(* IEC 61131-3 sources: 2026_Projet_YGO_ExcavatriceDragage/TOOLS/TEST_AUTO_CI/RESULTS/L_SIMULATION/tests (part 8) *)

TEST 'TC-T418-INT-004 Premier geste N2 observe HX1 existant'
nx := 5000; ny := 5000; raw1 := 0; raw2 := 0; previousButton := FALSE; buttonEdges := 0;
bench.Enable := TRUE; joy.Enable := TRUE; joy.ArmingPermit := TRUE; diagOk.Operational := TRUE;
joy.BusCanOpenOP := diagOk; joy.JoystickOP := diagOk; home.Enable := TRUE; home.BootReady := TRUE;
home.Mode := E_Mode.MAINT_N2; home.BucketOffsetValid := TRUE; home.WinchesMechanicallyStopped := TRUE;
ADVANCE_TIME(10000000);
bench(RawPosM1 := raw1, RawPosM2 := raw2);
joy(RawX := bench.Operator.JoyXRaw_ANA1, RawY := bench.Operator.JoyYRaw_ANA2, RawButton := bench.Operator.JoyBtnRaw, Cfg := cfg, NeutralXMem := nx, NeutralYMem := ny);
home(DeadmanArmed := joy.DeadmanArmed, JoystickDeflected := NOT joy.AtNeutralXY, JoystickPull := joy.AxisCmdY.DirectionPositive, JoystickPush := joy.AxisCmdY.DirectionNegative, BtnValidation := bench.Operator.JoyBtnRaw);
IF bench.Operator.JoyBtnRaw AND NOT previousButton THEN buttonEdges := buttonEdges + 1; END_IF; previousButton := bench.Operator.JoyBtnRaw;
bench.SimJoystickRight_Fwd_MAINT_Active := TRUE;
ADVANCE_TIME(10000000);
bench(RawPosM1 := raw1, RawPosM2 := raw2);
joy(RawX := bench.Operator.JoyXRaw_ANA1, RawY := bench.Operator.JoyYRaw_ANA2, RawButton := bench.Operator.JoyBtnRaw, Cfg := cfg, NeutralXMem := nx, NeutralYMem := ny);
home(DeadmanArmed := joy.DeadmanArmed, JoystickDeflected := NOT joy.AtNeutralXY, JoystickPull := joy.AxisCmdY.DirectionPositive, JoystickPush := joy.AxisCmdY.DirectionNegative, BtnValidation := bench.Operator.JoyBtnRaw);
IF bench.Operator.JoyBtnRaw AND NOT previousButton THEN buttonEdges := buttonEdges + 1; END_IF; previousButton := bench.Operator.JoyBtnRaw;
ASSERT_EQ(home.MachineHomingSeqStep, E_MachineHomingTxState.HX1_BUCKET_PREPARE, 'CONSTAT production : front homme-mort lance HX1 en N2');
ADVANCE_TIME(10000000);
bench(RawPosM1 := raw1, RawPosM2 := raw2);
joy(RawX := bench.Operator.JoyXRaw_ANA1, RawY := bench.Operator.JoyYRaw_ANA2, RawButton := bench.Operator.JoyBtnRaw, Cfg := cfg, NeutralXMem := nx, NeutralYMem := ny);
home(DeadmanArmed := joy.DeadmanArmed, JoystickDeflected := NOT joy.AtNeutralXY, JoystickPull := joy.AxisCmdY.DirectionPositive, JoystickPush := joy.AxisCmdY.DirectionNegative, BtnValidation := bench.Operator.JoyBtnRaw);
IF bench.Operator.JoyBtnRaw AND NOT previousButton THEN buttonEdges := buttonEdges + 1; END_IF; previousButton := bench.Operator.JoyBtnRaw;
ASSERT_TRUE(home.M3Locked, 'CONSTAT production : homing verrouille M3'); ASSERT_EQ(buttonEdges, 1, 'Front fidele non masque');
END_TEST

TEST 'TC-T418-INT-005 Stimuli manuels exclusifs et pas de saut au retour'
nx := 5000; ny := 5000; raw1 := 0; raw2 := 0; previousButton := FALSE; buttonEdges := 0;
bench.Enable := TRUE; joy.Enable := TRUE; joy.ArmingPermit := TRUE; diagOk.Operational := TRUE;
joy.BusCanOpenOP := diagOk; joy.JoystickOP := diagOk; home.Enable := TRUE; home.BootReady := TRUE;
home.Mode := E_Mode.MAINT_N1; home.BucketOffsetValid := TRUE; home.WinchesMechanicallyStopped := TRUE;
ADVANCE_TIME(10000000);
bench(RawPosM1 := raw1, RawPosM2 := raw2);
joy(RawX := bench.Operator.JoyXRaw_ANA1, RawY := bench.Operator.JoyYRaw_ANA2, RawButton := bench.Operator.JoyBtnRaw, Cfg := cfg, NeutralXMem := nx, NeutralYMem := ny);
home(DeadmanArmed := joy.DeadmanArmed, JoystickDeflected := NOT joy.AtNeutralXY, JoystickPull := joy.AxisCmdY.DirectionPositive, JoystickPush := joy.AxisCmdY.DirectionNegative, BtnValidation := bench.Operator.JoyBtnRaw);
IF bench.Operator.JoyBtnRaw AND NOT previousButton THEN buttonEdges := buttonEdges + 1; END_IF; previousButton := bench.Operator.JoyBtnRaw;
bench.SimJoystickRawX := 8000; bench.SimJoystickRawButton := TRUE;
ADVANCE_TIME(10000000);
bench(RawPosM1 := raw1, RawPosM2 := raw2);
joy(RawX := bench.Operator.JoyXRaw_ANA1, RawY := bench.Operator.JoyYRaw_ANA2, RawButton := bench.Operator.JoyBtnRaw, Cfg := cfg, NeutralXMem := nx, NeutralYMem := ny);
home(DeadmanArmed := joy.DeadmanArmed, JoystickDeflected := NOT joy.AtNeutralXY, JoystickPull := joy.AxisCmdY.DirectionPositive, JoystickPush := joy.AxisCmdY.DirectionNegative, BtnValidation := bench.Operator.JoyBtnRaw);
IF bench.Operator.JoyBtnRaw AND NOT previousButton THEN buttonEdges := buttonEdges + 1; END_IF; previousButton := bench.Operator.JoyBtnRaw;
ASSERT_EQ(bench.Operator.JoyXRaw_ANA1, 8000, 'Manuel disponible au repos'); ASSERT_TRUE(bench.Operator.JoyBtnRaw, 'Bouton manuel publie');
bench.SimJoystickRight_Fwd_MAINT_Active := TRUE;
ADVANCE_TIME(10000000);
bench(RawPosM1 := raw1, RawPosM2 := raw2);
joy(RawX := bench.Operator.JoyXRaw_ANA1, RawY := bench.Operator.JoyYRaw_ANA2, RawButton := bench.Operator.JoyBtnRaw, Cfg := cfg, NeutralXMem := nx, NeutralYMem := ny);
home(DeadmanArmed := joy.DeadmanArmed, JoystickDeflected := NOT joy.AtNeutralXY, JoystickPull := joy.AxisCmdY.DirectionPositive, JoystickPush := joy.AxisCmdY.DirectionNegative, BtnValidation := bench.Operator.JoyBtnRaw);
IF bench.Operator.JoyBtnRaw AND NOT previousButton THEN buttonEdges := buttonEdges + 1; END_IF; previousButton := bench.Operator.JoyBtnRaw;
ADVANCE_TIME(10000000);
bench(RawPosM1 := raw1, RawPosM2 := raw2);
joy(RawX := bench.Operator.JoyXRaw_ANA1, RawY := bench.Operator.JoyYRaw_ANA2, RawButton := bench.Operator.JoyBtnRaw, Cfg := cfg, NeutralXMem := nx, NeutralYMem := ny);
home(DeadmanArmed := joy.DeadmanArmed, JoystickDeflected := NOT joy.AtNeutralXY, JoystickPull := joy.AxisCmdY.DirectionPositive, JoystickPush := joy.AxisCmdY.DirectionNegative, BtnValidation := bench.Operator.JoyBtnRaw);
IF bench.Operator.JoyBtnRaw AND NOT previousButton THEN buttonEdges := buttonEdges + 1; END_IF; previousButton := bench.Operator.JoyBtnRaw;
ADVANCE_TIME(10000000);
bench(RawPosM1 := raw1, RawPosM2 := raw2);
joy(RawX := bench.Operator.JoyXRaw_ANA1, RawY := bench.Operator.JoyYRaw_ANA2, RawButton := bench.Operator.JoyBtnRaw, Cfg := cfg, NeutralXMem := nx, NeutralYMem := ny);
home(DeadmanArmed := joy.DeadmanArmed, JoystickDeflected := NOT joy.AtNeutralXY, JoystickPull := joy.AxisCmdY.DirectionPositive, JoystickPush := joy.AxisCmdY.DirectionNegative, BtnValidation := bench.Operator.JoyBtnRaw);
IF bench.Operator.JoyBtnRaw AND NOT previousButton THEN buttonEdges := buttonEdges + 1; END_IF; previousButton := bench.Operator.JoyBtnRaw;
ADVANCE_TIME(10000000);
bench(RawPosM1 := raw1, RawPosM2 := raw2);
joy(RawX := bench.Operator.JoyXRaw_ANA1, RawY := bench.Operator.JoyYRaw_ANA2, RawButton := bench.Operator.JoyBtnRaw, Cfg := cfg, NeutralXMem := nx, NeutralYMem := ny);
home(DeadmanArmed := joy.DeadmanArmed, JoystickDeflected := NOT joy.AtNeutralXY, JoystickPull := joy.AxisCmdY.DirectionPositive, JoystickPush := joy.AxisCmdY.DirectionNegative, BtnValidation := bench.Operator.JoyBtnRaw);
IF bench.Operator.JoyBtnRaw AND NOT previousButton THEN buttonEdges := buttonEdges + 1; END_IF; previousButton := bench.Operator.JoyBtnRaw;
ADVANCE_TIME(10000000);
bench(RawPosM1 := raw1, RawPosM2 := raw2);
joy(RawX := bench.Operator.JoyXRaw_ANA1, RawY := bench.Operator.JoyYRaw_ANA2, RawButton := bench.Operator.JoyBtnRaw, Cfg := cfg, NeutralXMem := nx, NeutralYMem := ny);
home(DeadmanArmed := joy.DeadmanArmed, JoystickDeflected := NOT joy.AtNeutralXY, JoystickPull := joy.AxisCmdY.DirectionPositive, JoystickPush := joy.AxisCmdY.DirectionNegative, BtnValidation := bench.Operator.JoyBtnRaw);
IF bench.Operator.JoyBtnRaw AND NOT previousButton THEN buttonEdges := buttonEdges + 1; END_IF; previousButton := bench.Operator.JoyBtnRaw;
ASSERT_EQ(bench.Operator.JoyXRaw_ANA1, 5000, 'Conflit manuel automatique neutralise'); ASSERT_FALSE(bench.Operator.JoyBtnRaw, 'Aucun OR des sources');
bench.SimJoystickRawX := 5000; bench.SimJoystickRawButton := FALSE;
ADVANCE_TIME(10000000);
bench(RawPosM1 := raw1, RawPosM2 := raw2);
joy(RawX := bench.Operator.JoyXRaw_ANA1, RawY := bench.Operator.JoyYRaw_ANA2, RawButton := bench.Operator.JoyBtnRaw, Cfg := cfg, NeutralXMem := nx, NeutralYMem := ny);
home(DeadmanArmed := joy.DeadmanArmed, JoystickDeflected := NOT joy.AtNeutralXY, JoystickPull := joy.AxisCmdY.DirectionPositive, JoystickPush := joy.AxisCmdY.DirectionNegative, BtnValidation := bench.Operator.JoyBtnRaw);
IF bench.Operator.JoyBtnRaw AND NOT previousButton THEN buttonEdges := buttonEdges + 1; END_IF; previousButton := bench.Operator.JoyBtnRaw;
ADVANCE_TIME(10000000);
bench(RawPosM1 := raw1, RawPosM2 := raw2);
joy(RawX := bench.Operator.JoyXRaw_ANA1, RawY := bench.Operator.JoyYRaw_ANA2, RawButton := bench.Operator.JoyBtnRaw, Cfg := cfg, NeutralXMem := nx, NeutralYMem := ny);
home(DeadmanArmed := joy.DeadmanArmed, JoystickDeflected := NOT joy.AtNeutralXY, JoystickPull := joy.AxisCmdY.DirectionPositive, JoystickPush := joy.AxisCmdY.DirectionNegative, BtnValidation := bench.Operator.JoyBtnRaw);
IF bench.Operator.JoyBtnRaw AND NOT previousButton THEN buttonEdges := buttonEdges + 1; END_IF; previousButton := bench.Operator.JoyBtnRaw;
ADVANCE_TIME(10000000);
bench(RawPosM1 := raw1, RawPosM2 := raw2);
joy(RawX := bench.Operator.JoyXRaw_ANA1, RawY := bench.Operator.JoyYRaw_ANA2, RawButton := bench.Operator.JoyBtnRaw, Cfg := cfg, NeutralXMem := nx, NeutralYMem := ny);
home(DeadmanArmed := joy.DeadmanArmed, JoystickDeflected := NOT joy.AtNeutralXY, JoystickPull := joy.AxisCmdY.DirectionPositive, JoystickPush := joy.AxisCmdY.DirectionNegative, BtnValidation := bench.Operator.JoyBtnRaw);
IF bench.Operator.JoyBtnRaw AND NOT previousButton THEN buttonEdges := buttonEdges + 1; END_IF; previousButton := bench.Operator.JoyBtnRaw;
ADVANCE_TIME(10000000);
bench(RawPosM1 := raw1, RawPosM2 := raw2);
joy(RawX := bench.Operator.JoyXRaw_ANA1, RawY := bench.Operator.JoyYRaw_ANA2, RawButton := bench.Operator.JoyBtnRaw, Cfg := cfg, NeutralXMem := nx, NeutralYMem := ny);
home(DeadmanArmed := joy.DeadmanArmed, JoystickDeflected := NOT joy.AtNeutralXY, JoystickPull := joy.AxisCmdY.DirectionPositive, JoystickPush := joy.AxisCmdY.DirectionNegative, BtnValidation := bench.Operator.JoyBtnRaw);
IF bench.Operator.JoyBtnRaw AND NOT previousButton THEN buttonEdges := buttonEdges + 1; END_IF; previousButton := bench.Operator.JoyBtnRaw;
ADVANCE_TIME(10000000);
bench(RawPosM1 := raw1, RawPosM2 := raw2);
joy(RawX := bench.Operator.JoyXRaw_ANA1, RawY := bench.Operator.JoyYRaw_ANA2, RawButton := bench.Operator.JoyBtnRaw, Cfg := cfg, NeutralXMem := nx, NeutralYMem := ny);
home(DeadmanArmed := joy.DeadmanArmed, JoystickDeflected := NOT joy.AtNeutralXY, JoystickPull := joy.AxisCmdY.DirectionPositive, JoystickPush := joy.AxisCmdY.DirectionNegative, BtnValidation := bench.Operator.JoyBtnRaw);
IF bench.Operator.JoyBtnRaw AND NOT previousButton THEN buttonEdges := buttonEdges + 1; END_IF; previousButton := bench.Operator.JoyBtnRaw;
ASSERT_FALSE(bench.Operator.JoyBtnRaw, 'Enlever stimulus ne demarre pas bouton tenu');
bench.SimJoystickRight_Fwd_MAINT_Active := FALSE;
ADVANCE_TIME(10000000);
bench(RawPosM1 := raw1, RawPosM2 := raw2);
joy(RawX := bench.Operator.JoyXRaw_ANA1, RawY := bench.Operator.JoyYRaw_ANA2, RawButton := bench.Operator.JoyBtnRaw, Cfg := cfg, NeutralXMem := nx, NeutralYMem := ny);
home(DeadmanArmed := joy.DeadmanArmed, JoystickDeflected := NOT joy.AtNeutralXY, JoystickPull := joy.AxisCmdY.DirectionPositive, JoystickPush := joy.AxisCmdY.DirectionNegative, BtnValidation := bench.Operator.JoyBtnRaw);
IF bench.Operator.JoyBtnRaw AND NOT previousButton THEN buttonEdges := buttonEdges + 1; END_IF; previousButton := bench.Operator.JoyBtnRaw;
bench.SimJoystickRight_Fwd_MAINT_Active := TRUE;
ADVANCE_TIME(10000000);
bench(RawPosM1 := raw1, RawPosM2 := raw2);
joy(RawX := bench.Operator.JoyXRaw_ANA1, RawY := bench.Operator.JoyYRaw_ANA2, RawButton := bench.Operator.JoyBtnRaw, Cfg := cfg, NeutralXMem := nx, NeutralYMem := ny);
home(DeadmanArmed := joy.DeadmanArmed, JoystickDeflected := NOT joy.AtNeutralXY, JoystickPull := joy.AxisCmdY.DirectionPositive, JoystickPush := joy.AxisCmdY.DirectionNegative, BtnValidation := bench.Operator.JoyBtnRaw);
IF bench.Operator.JoyBtnRaw AND NOT previousButton THEN buttonEdges := buttonEdges + 1; END_IF; previousButton := bench.Operator.JoyBtnRaw;
ADVANCE_TIME(10000000);
bench(RawPosM1 := raw1, RawPosM2 := raw2);
joy(RawX := bench.Operator.JoyXRaw_ANA1, RawY := bench.Operator.JoyYRaw_ANA2, RawButton := bench.Operator.JoyBtnRaw, Cfg := cfg, NeutralXMem := nx, NeutralYMem := ny);
home(DeadmanArmed := joy.DeadmanArmed, JoystickDeflected := NOT joy.AtNeutralXY, JoystickPull := joy.AxisCmdY.DirectionPositive, JoystickPush := joy.AxisCmdY.DirectionNegative, BtnValidation := bench.Operator.JoyBtnRaw);
IF bench.Operator.JoyBtnRaw AND NOT previousButton THEN buttonEdges := buttonEdges + 1; END_IF; previousButton := bench.Operator.JoyBtnRaw;
ADVANCE_TIME(10000000);
bench(RawPosM1 := raw1, RawPosM2 := raw2);
joy(RawX := bench.Operator.JoyXRaw_ANA1, RawY := bench.Operator.JoyYRaw_ANA2, RawButton := bench.Operator.JoyBtnRaw, Cfg := cfg, NeutralXMem := nx, NeutralYMem := ny);
home(DeadmanArmed := joy.DeadmanArmed, JoystickDeflected := NOT joy.AtNeutralXY, JoystickPull := joy.AxisCmdY.DirectionPositive, JoystickPush := joy.AxisCmdY.DirectionNegative, BtnValidation := bench.Operator.JoyBtnRaw);
IF bench.Operator.JoyBtnRaw AND NOT previousButton THEN buttonEdges := buttonEdges + 1; END_IF; previousButton := bench.Operator.JoyBtnRaw;
ADVANCE_TIME(10000000);
bench(RawPosM1 := raw1, RawPosM2 := raw2);
joy(RawX := bench.Operator.JoyXRaw_ANA1, RawY := bench.Operator.JoyYRaw_ANA2, RawButton := bench.Operator.JoyBtnRaw, Cfg := cfg, NeutralXMem := nx, NeutralYMem := ny);
home(DeadmanArmed := joy.DeadmanArmed, JoystickDeflected := NOT joy.AtNeutralXY, JoystickPull := joy.AxisCmdY.DirectionPositive, JoystickPush := joy.AxisCmdY.DirectionNegative, BtnValidation := bench.Operator.JoyBtnRaw);
IF bench.Operator.JoyBtnRaw AND NOT previousButton THEN buttonEdges := buttonEdges + 1; END_IF; previousButton := bench.Operator.JoyBtnRaw;
ADVANCE_TIME(10000000);
bench(RawPosM1 := raw1, RawPosM2 := raw2);
joy(RawX := bench.Operator.JoyXRaw_ANA1, RawY := bench.Operator.JoyYRaw_ANA2, RawButton := bench.Operator.JoyBtnRaw, Cfg := cfg, NeutralXMem := nx, NeutralYMem := ny);
home(DeadmanArmed := joy.DeadmanArmed, JoystickDeflected := NOT joy.AtNeutralXY, JoystickPull := joy.AxisCmdY.DirectionPositive, JoystickPush := joy.AxisCmdY.DirectionNegative, BtnValidation := bench.Operator.JoyBtnRaw);
IF bench.Operator.JoyBtnRaw AND NOT previousButton THEN buttonEdges := buttonEdges + 1; END_IF; previousButton := bench.Operator.JoyBtnRaw;
ADVANCE_TIME(10000000);
bench(RawPosM1 := raw1, RawPosM2 := raw2);
joy(RawX := bench.Operator.JoyXRaw_ANA1, RawY := bench.Operator.JoyYRaw_ANA2, RawButton := bench.Operator.JoyBtnRaw, Cfg := cfg, NeutralXMem := nx, NeutralYMem := ny);
home(DeadmanArmed := joy.DeadmanArmed, JoystickDeflected := NOT joy.AtNeutralXY, JoystickPull := joy.AxisCmdY.DirectionPositive, JoystickPush := joy.AxisCmdY.DirectionNegative, BtnValidation := bench.Operator.JoyBtnRaw);
IF bench.Operator.JoyBtnRaw AND NOT previousButton THEN buttonEdges := buttonEdges + 1; END_IF; previousButton := bench.Operator.JoyBtnRaw;
ADVANCE_TIME(10000000);
bench(RawPosM1 := raw1, RawPosM2 := raw2);
joy(RawX := bench.Operator.JoyXRaw_ANA1, RawY := bench.Operator.JoyYRaw_ANA2, RawButton := bench.Operator.JoyBtnRaw, Cfg := cfg, NeutralXMem := nx, NeutralYMem := ny);
home(DeadmanArmed := joy.DeadmanArmed, JoystickDeflected := NOT joy.AtNeutralXY, JoystickPull := joy.AxisCmdY.DirectionPositive, JoystickPush := joy.AxisCmdY.DirectionNegative, BtnValidation := bench.Operator.JoyBtnRaw);
IF bench.Operator.JoyBtnRaw AND NOT previousButton THEN buttonEdges := buttonEdges + 1; END_IF; previousButton := bench.Operator.JoyBtnRaw;
ADVANCE_TIME(10000000);
bench(RawPosM1 := raw1, RawPosM2 := raw2);
joy(RawX := bench.Operator.JoyXRaw_ANA1, RawY := bench.Operator.JoyYRaw_ANA2, RawButton := bench.Operator.JoyBtnRaw, Cfg := cfg, NeutralXMem := nx, NeutralYMem := ny);
home(DeadmanArmed := joy.DeadmanArmed, JoystickDeflected := NOT joy.AtNeutralXY, JoystickPull := joy.AxisCmdY.DirectionPositive, JoystickPush := joy.AxisCmdY.DirectionNegative, BtnValidation := bench.Operator.JoyBtnRaw);
IF bench.Operator.JoyBtnRaw AND NOT previousButton THEN buttonEdges := buttonEdges + 1; END_IF; previousButton := bench.Operator.JoyBtnRaw;
ADVANCE_TIME(10000000);
bench(RawPosM1 := raw1, RawPosM2 := raw2);
joy(RawX := bench.Operator.JoyXRaw_ANA1, RawY := bench.Operator.JoyYRaw_ANA2, RawButton := bench.Operator.JoyBtnRaw, Cfg := cfg, NeutralXMem := nx, NeutralYMem := ny);
home(DeadmanArmed := joy.DeadmanArmed, JoystickDeflected := NOT joy.AtNeutralXY, JoystickPull := joy.AxisCmdY.DirectionPositive, JoystickPush := joy.AxisCmdY.DirectionNegative, BtnValidation := bench.Operator.JoyBtnRaw);
IF bench.Operator.JoyBtnRaw AND NOT previousButton THEN buttonEdges := buttonEdges + 1; END_IF; previousButton := bench.Operator.JoyBtnRaw;
ADVANCE_TIME(10000000);
bench(RawPosM1 := raw1, RawPosM2 := raw2);
joy(RawX := bench.Operator.JoyXRaw_ANA1, RawY := bench.Operator.JoyYRaw_ANA2, RawButton := bench.Operator.JoyBtnRaw, Cfg := cfg, NeutralXMem := nx, NeutralYMem := ny);
home(DeadmanArmed := joy.DeadmanArmed, JoystickDeflected := NOT joy.AtNeutralXY, JoystickPull := joy.AxisCmdY.DirectionPositive, JoystickPush := joy.AxisCmdY.DirectionNegative, BtnValidation := bench.Operator.JoyBtnRaw);
IF bench.Operator.JoyBtnRaw AND NOT previousButton THEN buttonEdges := buttonEdges + 1; END_IF; previousButton := bench.Operator.JoyBtnRaw;
ADVANCE_TIME(10000000);
bench(RawPosM1 := raw1, RawPosM2 := raw2);
joy(RawX := bench.Operator.JoyXRaw_ANA1, RawY := bench.Operator.JoyYRaw_ANA2, RawButton := bench.Operator.JoyBtnRaw, Cfg := cfg, NeutralXMem := nx, NeutralYMem := ny);
home(DeadmanArmed := joy.DeadmanArmed, JoystickDeflected := NOT joy.AtNeutralXY, JoystickPull := joy.AxisCmdY.DirectionPositive, JoystickPush := joy.AxisCmdY.DirectionNegative, BtnValidation := bench.Operator.JoyBtnRaw);
IF bench.Operator.JoyBtnRaw AND NOT previousButton THEN buttonEdges := buttonEdges + 1; END_IF; previousButton := bench.Operator.JoyBtnRaw;
ADVANCE_TIME(10000000);
bench(RawPosM1 := raw1, RawPosM2 := raw2);
joy(RawX := bench.Operator.JoyXRaw_ANA1, RawY := bench.Operator.JoyYRaw_ANA2, RawButton := bench.Operator.JoyBtnRaw, Cfg := cfg, NeutralXMem := nx, NeutralYMem := ny);
home(DeadmanArmed := joy.DeadmanArmed, JoystickDeflected := NOT joy.AtNeutralXY, JoystickPull := joy.AxisCmdY.DirectionPositive, JoystickPush := joy.AxisCmdY.DirectionNegative, BtnValidation := bench.Operator.JoyBtnRaw);
IF bench.Operator.JoyBtnRaw AND NOT previousButton THEN buttonEdges := buttonEdges + 1; END_IF; previousButton := bench.Operator.JoyBtnRaw;
ADVANCE_TIME(10000000);
bench(RawPosM1 := raw1, RawPosM2 := raw2);
joy(RawX := bench.Operator.JoyXRaw_ANA1, RawY := bench.Operator.JoyYRaw_ANA2, RawButton := bench.Operator.JoyBtnRaw, Cfg := cfg, NeutralXMem := nx, NeutralYMem := ny);
home(DeadmanArmed := joy.DeadmanArmed, JoystickDeflected := NOT joy.AtNeutralXY, JoystickPull := joy.AxisCmdY.DirectionPositive, JoystickPush := joy.AxisCmdY.DirectionNegative, BtnValidation := bench.Operator.JoyBtnRaw);
IF bench.Operator.JoyBtnRaw AND NOT previousButton THEN buttonEdges := buttonEdges + 1; END_IF; previousButton := bench.Operator.JoyBtnRaw;
ADVANCE_TIME(10000000);
bench(RawPosM1 := raw1, RawPosM2 := raw2);
joy(RawX := bench.Operator.JoyXRaw_ANA1, RawY := bench.Operator.JoyYRaw_ANA2, RawButton := bench.Operator.JoyBtnRaw, Cfg := cfg, NeutralXMem := nx, NeutralYMem := ny);
home(DeadmanArmed := joy.DeadmanArmed, JoystickDeflected := NOT joy.AtNeutralXY, JoystickPull := joy.AxisCmdY.DirectionPositive, JoystickPush := joy.AxisCmdY.DirectionNegative, BtnValidation := bench.Operator.JoyBtnRaw);
IF bench.Operator.JoyBtnRaw AND NOT previousButton THEN buttonEdges := buttonEdges + 1; END_IF; previousButton := bench.Operator.JoyBtnRaw;
ADVANCE_TIME(10000000);
bench(RawPosM1 := raw1, RawPosM2 := raw2);
joy(RawX := bench.Operator.JoyXRaw_ANA1, RawY := bench.Operator.JoyYRaw_ANA2, RawButton := bench.Operator.JoyBtnRaw, Cfg := cfg, NeutralXMem := nx, NeutralYMem := ny);
home(DeadmanArmed := joy.DeadmanArmed, JoystickDeflected := NOT joy.AtNeutralXY, JoystickPull := joy.AxisCmdY.DirectionPositive, JoystickPush := joy.AxisCmdY.DirectionNegative, BtnValidation := bench.Operator.JoyBtnRaw);
IF bench.Operator.JoyBtnRaw AND NOT previousButton THEN buttonEdges := buttonEdges + 1; END_IF; previousButton := bench.Operator.JoyBtnRaw;
ADVANCE_TIME(10000000);
bench(RawPosM1 := raw1, RawPosM2 := raw2);
joy(RawX := bench.Operator.JoyXRaw_ANA1, RawY := bench.Operator.JoyYRaw_ANA2, RawButton := bench.Operator.JoyBtnRaw, Cfg := cfg, NeutralXMem := nx, NeutralYMem := ny);
home(DeadmanArmed := joy.DeadmanArmed, JoystickDeflected := NOT joy.AtNeutralXY, JoystickPull := joy.AxisCmdY.DirectionPositive, JoystickPush := joy.AxisCmdY.DirectionNegative, BtnValidation := bench.Operator.JoyBtnRaw);
IF bench.Operator.JoyBtnRaw AND NOT previousButton THEN buttonEdges := buttonEdges + 1; END_IF; previousButton := bench.Operator.JoyBtnRaw;
ADVANCE_TIME(10000000);
bench(RawPosM1 := raw1, RawPosM2 := raw2);
joy(RawX := bench.Operator.JoyXRaw_ANA1, RawY := bench.Operator.JoyYRaw_ANA2, RawButton := bench.Operator.JoyBtnRaw, Cfg := cfg, NeutralXMem := nx, NeutralYMem := ny);
home(DeadmanArmed := joy.DeadmanArmed, JoystickDeflected := NOT joy.AtNeutralXY, JoystickPull := joy.AxisCmdY.DirectionPositive, JoystickPush := joy.AxisCmdY.DirectionNegative, BtnValidation := bench.Operator.JoyBtnRaw);
IF bench.Operator.JoyBtnRaw AND NOT previousButton THEN buttonEdges := buttonEdges + 1; END_IF; previousButton := bench.Operator.JoyBtnRaw;
ADVANCE_TIME(10000000);
bench(RawPosM1 := raw1, RawPosM2 := raw2);
joy(RawX := bench.Operator.JoyXRaw_ANA1, RawY := bench.Operator.JoyYRaw_ANA2, RawButton := bench.Operator.JoyBtnRaw, Cfg := cfg, NeutralXMem := nx, NeutralYMem := ny);
home(DeadmanArmed := joy.DeadmanArmed, JoystickDeflected := NOT joy.AtNeutralXY, JoystickPull := joy.AxisCmdY.DirectionPositive, JoystickPush := joy.AxisCmdY.DirectionNegative, BtnValidation := bench.Operator.JoyBtnRaw);
IF bench.Operator.JoyBtnRaw AND NOT previousButton THEN buttonEdges := buttonEdges + 1; END_IF; previousButton := bench.Operator.JoyBtnRaw;
ADVANCE_TIME(10000000);
bench(RawPosM1 := raw1, RawPosM2 := raw2);
joy(RawX := bench.Operator.JoyXRaw_ANA1, RawY := bench.Operator.JoyYRaw_ANA2, RawButton := bench.Operator.JoyBtnRaw, Cfg := cfg, NeutralXMem := nx, NeutralYMem := ny);
home(DeadmanArmed := joy.DeadmanArmed, JoystickDeflected := NOT joy.AtNeutralXY, JoystickPull := joy.AxisCmdY.DirectionPositive, JoystickPush := joy.AxisCmdY.DirectionNegative, BtnValidation := bench.Operator.JoyBtnRaw);
IF bench.Operator.JoyBtnRaw AND NOT previousButton THEN buttonEdges := buttonEdges + 1; END_IF; previousButton := bench.Operator.JoyBtnRaw;
ADVANCE_TIME(10000000);
bench(RawPosM1 := raw1, RawPosM2 := raw2);
joy(RawX := bench.Operator.JoyXRaw_ANA1, RawY := bench.Operator.JoyYRaw_ANA2, RawButton := bench.Operator.JoyBtnRaw, Cfg := cfg, NeutralXMem := nx, NeutralYMem := ny);
home(DeadmanArmed := joy.DeadmanArmed, JoystickDeflected := NOT joy.AtNeutralXY, JoystickPull := joy.AxisCmdY.DirectionPositive, JoystickPush := joy.AxisCmdY.DirectionNegative, BtnValidation := bench.Operator.JoyBtnRaw);
IF bench.Operator.JoyBtnRaw AND NOT previousButton THEN buttonEdges := buttonEdges + 1; END_IF; previousButton := bench.Operator.JoyBtnRaw;
ADVANCE_TIME(10000000);
bench(RawPosM1 := raw1, RawPosM2 := raw2);
joy(RawX := bench.Operator.JoyXRaw_ANA1, RawY := bench.Operator.JoyYRaw_ANA2, RawButton := bench.Operator.JoyBtnRaw, Cfg := cfg, NeutralXMem := nx, NeutralYMem := ny);
home(DeadmanArmed := joy.DeadmanArmed, JoystickDeflected := NOT joy.AtNeutralXY, JoystickPull := joy.AxisCmdY.DirectionPositive, JoystickPush := joy.AxisCmdY.DirectionNegative, BtnValidation := bench.Operator.JoyBtnRaw);
IF bench.Operator.JoyBtnRaw AND NOT previousButton THEN buttonEdges := buttonEdges + 1; END_IF; previousButton := bench.Operator.JoyBtnRaw;
ADVANCE_TIME(10000000);
bench(RawPosM1 := raw1, RawPosM2 := raw2);
joy(RawX := bench.Operator.JoyXRaw_ANA1, RawY := bench.Operator.JoyYRaw_ANA2, RawButton := bench.Operator.JoyBtnRaw, Cfg := cfg, NeutralXMem := nx, NeutralYMem := ny);
home(DeadmanArmed := joy.DeadmanArmed, JoystickDeflected := NOT joy.AtNeutralXY, JoystickPull := joy.AxisCmdY.DirectionPositive, JoystickPush := joy.AxisCmdY.DirectionNegative, BtnValidation := bench.Operator.JoyBtnRaw);
IF bench.Operator.JoyBtnRaw AND NOT previousButton THEN buttonEdges := buttonEdges + 1; END_IF; previousButton := bench.Operator.JoyBtnRaw;
ADVANCE_TIME(10000000);
bench(RawPosM1 := raw1, RawPosM2 := raw2);
joy(RawX := bench.Operator.JoyXRaw_ANA1, RawY := bench.Operator.JoyYRaw_ANA2, RawButton := bench.Operator.JoyBtnRaw, Cfg := cfg, NeutralXMem := nx, NeutralYMem := ny);
home(DeadmanArmed := joy.DeadmanArmed, JoystickDeflected := NOT joy.AtNeutralXY, JoystickPull := joy.AxisCmdY.DirectionPositive, JoystickPush := joy.AxisCmdY.DirectionNegative, BtnValidation := bench.Operator.JoyBtnRaw);
IF bench.Operator.JoyBtnRaw AND NOT previousButton THEN buttonEdges := buttonEdges + 1; END_IF; previousButton := bench.Operator.JoyBtnRaw;
ADVANCE_TIME(10000000);
bench(RawPosM1 := raw1, RawPosM2 := raw2);
joy(RawX := bench.Operator.JoyXRaw_ANA1, RawY := bench.Operator.JoyYRaw_ANA2, RawButton := bench.Operator.JoyBtnRaw, Cfg := cfg, NeutralXMem := nx, NeutralYMem := ny);
home(DeadmanArmed := joy.DeadmanArmed, JoystickDeflected := NOT joy.AtNeutralXY, JoystickPull := joy.AxisCmdY.DirectionPositive, JoystickPush := joy.AxisCmdY.DirectionNegative, BtnValidation := bench.Operator.JoyBtnRaw);
IF bench.Operator.JoyBtnRaw AND NOT previousButton THEN buttonEdges := buttonEdges + 1; END_IF; previousButton := bench.Operator.JoyBtnRaw;
ADVANCE_TIME(10000000);
bench(RawPosM1 := raw1, RawPosM2 := raw2);
joy(RawX := bench.Operator.JoyXRaw_ANA1, RawY := bench.Operator.JoyYRaw_ANA2, RawButton := bench.Operator.JoyBtnRaw, Cfg := cfg, NeutralXMem := nx, NeutralYMem := ny);
home(DeadmanArmed := joy.DeadmanArmed, JoystickDeflected := NOT joy.AtNeutralXY, JoystickPull := joy.AxisCmdY.DirectionPositive, JoystickPush := joy.AxisCmdY.DirectionNegative, BtnValidation := bench.Operator.JoyBtnRaw);
IF bench.Operator.JoyBtnRaw AND NOT previousButton THEN buttonEdges := buttonEdges + 1; END_IF; previousButton := bench.Operator.JoyBtnRaw;
ADVANCE_TIME(10000000);
bench(RawPosM1 := raw1, RawPosM2 := raw2);
joy(RawX := bench.Operator.JoyXRaw_ANA1, RawY := bench.Operator.JoyYRaw_ANA2, RawButton := bench.Operator.JoyBtnRaw, Cfg := cfg, NeutralXMem := nx, NeutralYMem := ny);
home(DeadmanArmed := joy.DeadmanArmed, JoystickDeflected := NOT joy.AtNeutralXY, JoystickPull := joy.AxisCmdY.DirectionPositive, JoystickPush := joy.AxisCmdY.DirectionNegative, BtnValidation := bench.Operator.JoyBtnRaw);
IF bench.Operator.JoyBtnRaw AND NOT previousButton THEN buttonEdges := buttonEdges + 1; END_IF; previousButton := bench.Operator.JoyBtnRaw;
ADVANCE_TIME(10000000);
bench(RawPosM1 := raw1, RawPosM2 := raw2);
joy(RawX := bench.Operator.JoyXRaw_ANA1, RawY := bench.Operator.JoyYRaw_ANA2, RawButton := bench.Operator.JoyBtnRaw, Cfg := cfg, NeutralXMem := nx, NeutralYMem := ny);
home(DeadmanArmed := joy.DeadmanArmed, JoystickDeflected := NOT joy.AtNeutralXY, JoystickPull := joy.AxisCmdY.DirectionPositive, JoystickPush := joy.AxisCmdY.DirectionNegative, BtnValidation := bench.Operator.JoyBtnRaw);
IF bench.Operator.JoyBtnRaw AND NOT previousButton THEN buttonEdges := buttonEdges + 1; END_IF; previousButton := bench.Operator.JoyBtnRaw;
ADVANCE_TIME(10000000);
bench(RawPosM1 := raw1, RawPosM2 := raw2);
joy(RawX := bench.Operator.JoyXRaw_ANA1, RawY := bench.Operator.JoyYRaw_ANA2, RawButton := bench.Operator.JoyBtnRaw, Cfg := cfg, NeutralXMem := nx, NeutralYMem := ny);
home(DeadmanArmed := joy.DeadmanArmed, JoystickDeflected := NOT joy.AtNeutralXY, JoystickPull := joy.AxisCmdY.DirectionPositive, JoystickPush := joy.AxisCmdY.DirectionNegative, BtnValidation := bench.Operator.JoyBtnRaw);
IF bench.Operator.JoyBtnRaw AND NOT previousButton THEN buttonEdges := buttonEdges + 1; END_IF; previousButton := bench.Operator.JoyBtnRaw;
ADVANCE_TIME(10000000);
bench(RawPosM1 := raw1, RawPosM2 := raw2);
joy(RawX := bench.Operator.JoyXRaw_ANA1, RawY := bench.Operator.JoyYRaw_ANA2, RawButton := bench.Operator.JoyBtnRaw, Cfg := cfg, NeutralXMem := nx, NeutralYMem := ny);
home(DeadmanArmed := joy.DeadmanArmed, JoystickDeflected := NOT joy.AtNeutralXY, JoystickPull := joy.AxisCmdY.DirectionPositive, JoystickPush := joy.AxisCmdY.DirectionNegative, BtnValidation := bench.Operator.JoyBtnRaw);
IF bench.Operator.JoyBtnRaw AND NOT previousButton THEN buttonEdges := buttonEdges + 1; END_IF; previousButton := bench.Operator.JoyBtnRaw;
ADVANCE_TIME(10000000);
bench(RawPosM1 := raw1, RawPosM2 := raw2);
joy(RawX := bench.Operator.JoyXRaw_ANA1, RawY := bench.Operator.JoyYRaw_ANA2, RawButton := bench.Operator.JoyBtnRaw, Cfg := cfg, NeutralXMem := nx, NeutralYMem := ny);
home(DeadmanArmed := joy.DeadmanArmed, JoystickDeflected := NOT joy.AtNeutralXY, JoystickPull := joy.AxisCmdY.DirectionPositive, JoystickPush := joy.AxisCmdY.DirectionNegative, BtnValidation := bench.Operator.JoyBtnRaw);
IF bench.Operator.JoyBtnRaw AND NOT previousButton THEN buttonEdges := buttonEdges + 1; END_IF; previousButton := bench.Operator.JoyBtnRaw;
ADVANCE_TIME(10000000);
bench(RawPosM1 := raw1, RawPosM2 := raw2);
joy(RawX := bench.Operator.JoyXRaw_ANA1, RawY := bench.Operator.JoyYRaw_ANA2, RawButton := bench.Operator.JoyBtnRaw, Cfg := cfg, NeutralXMem := nx, NeutralYMem := ny);
home(DeadmanArmed := joy.DeadmanArmed, JoystickDeflected := NOT joy.AtNeutralXY, JoystickPull := joy.AxisCmdY.DirectionPositive, JoystickPush := joy.AxisCmdY.DirectionNegative, BtnValidation := bench.Operator.JoyBtnRaw);
IF bench.Operator.JoyBtnRaw AND NOT previousButton THEN buttonEdges := buttonEdges + 1; END_IF; previousButton := bench.Operator.JoyBtnRaw;
ADVANCE_TIME(10000000);
bench(RawPosM1 := raw1, RawPosM2 := raw2);
joy(RawX := bench.Operator.JoyXRaw_ANA1, RawY := bench.Operator.JoyYRaw_ANA2, RawButton := bench.Operator.JoyBtnRaw, Cfg := cfg, NeutralXMem := nx, NeutralYMem := ny);
home(DeadmanArmed := joy.DeadmanArmed, JoystickDeflected := NOT joy.AtNeutralXY, JoystickPull := joy.AxisCmdY.DirectionPositive, JoystickPush := joy.AxisCmdY.DirectionNegative, BtnValidation := bench.Operator.JoyBtnRaw);
IF bench.Operator.JoyBtnRaw AND NOT previousButton THEN buttonEdges := buttonEdges + 1; END_IF; previousButton := bench.Operator.JoyBtnRaw;
ADVANCE_TIME(10000000);
bench(RawPosM1 := raw1, RawPosM2 := raw2);
joy(RawX := bench.Operator.JoyXRaw_ANA1, RawY := bench.Operator.JoyYRaw_ANA2, RawButton := bench.Operator.JoyBtnRaw, Cfg := cfg, NeutralXMem := nx, NeutralYMem := ny);
home(DeadmanArmed := joy.DeadmanArmed, JoystickDeflected := NOT joy.AtNeutralXY, JoystickPull := joy.AxisCmdY.DirectionPositive, JoystickPush := joy.AxisCmdY.DirectionNegative, BtnValidation := bench.Operator.JoyBtnRaw);
IF bench.Operator.JoyBtnRaw AND NOT previousButton THEN buttonEdges := buttonEdges + 1; END_IF; previousButton := bench.Operator.JoyBtnRaw;
ADVANCE_TIME(10000000);
bench(RawPosM1 := raw1, RawPosM2 := raw2);
joy(RawX := bench.Operator.JoyXRaw_ANA1, RawY := bench.Operator.JoyYRaw_ANA2, RawButton := bench.Operator.JoyBtnRaw, Cfg := cfg, NeutralXMem := nx, NeutralYMem := ny);
home(DeadmanArmed := joy.DeadmanArmed, JoystickDeflected := NOT joy.AtNeutralXY, JoystickPull := joy.AxisCmdY.DirectionPositive, JoystickPush := joy.AxisCmdY.DirectionNegative, BtnValidation := bench.Operator.JoyBtnRaw);
IF bench.Operator.JoyBtnRaw AND NOT previousButton THEN buttonEdges := buttonEdges + 1; END_IF; previousButton := bench.Operator.JoyBtnRaw;
ADVANCE_TIME(10000000);
bench(RawPosM1 := raw1, RawPosM2 := raw2);
joy(RawX := bench.Operator.JoyXRaw_ANA1, RawY := bench.Operator.JoyYRaw_ANA2, RawButton := bench.Operator.JoyBtnRaw, Cfg := cfg, NeutralXMem := nx, NeutralYMem := ny);
home(DeadmanArmed := joy.DeadmanArmed, JoystickDeflected := NOT joy.AtNeutralXY, JoystickPull := joy.AxisCmdY.DirectionPositive, JoystickPush := joy.AxisCmdY.DirectionNegative, BtnValidation := bench.Operator.JoyBtnRaw);
IF bench.Operator.JoyBtnRaw AND NOT previousButton THEN buttonEdges := buttonEdges + 1; END_IF; previousButton := bench.Operator.JoyBtnRaw;
ADVANCE_TIME(10000000);
bench(RawPosM1 := raw1, RawPosM2 := raw2);
joy(RawX := bench.Operator.JoyXRaw_ANA1, RawY := bench.Operator.JoyYRaw_ANA2, RawButton := bench.Operator.JoyBtnRaw, Cfg := cfg, NeutralXMem := nx, NeutralYMem := ny);
home(DeadmanArmed := joy.DeadmanArmed, JoystickDeflected := NOT joy.AtNeutralXY, JoystickPull := joy.AxisCmdY.DirectionPositive, JoystickPush := joy.AxisCmdY.DirectionNegative, BtnValidation := bench.Operator.JoyBtnRaw);
IF bench.Operator.JoyBtnRaw AND NOT previousButton THEN buttonEdges := buttonEdges + 1; END_IF; previousButton := bench.Operator.JoyBtnRaw;
ADVANCE_TIME(10000000);
bench(RawPosM1 := raw1, RawPosM2 := raw2);
joy(RawX := bench.Operator.JoyXRaw_ANA1, RawY := bench.Operator.JoyYRaw_ANA2, RawButton := bench.Operator.JoyBtnRaw, Cfg := cfg, NeutralXMem := nx, NeutralYMem := ny);
home(DeadmanArmed := joy.DeadmanArmed, JoystickDeflected := NOT joy.AtNeutralXY, JoystickPull := joy.AxisCmdY.DirectionPositive, JoystickPush := joy.AxisCmdY.DirectionNegative, BtnValidation := bench.Operator.JoyBtnRaw);
IF bench.Operator.JoyBtnRaw AND NOT previousButton THEN buttonEdges := buttonEdges + 1; END_IF; previousButton := bench.Operator.JoyBtnRaw;
ADVANCE_TIME(10000000);
bench(RawPosM1 := raw1, RawPosM2 := raw2);
joy(RawX := bench.Operator.JoyXRaw_ANA1, RawY := bench.Operator.JoyYRaw_ANA2, RawButton := bench.Operator.JoyBtnRaw, Cfg := cfg, NeutralXMem := nx, NeutralYMem := ny);
home(DeadmanArmed := joy.DeadmanArmed, JoystickDeflected := NOT joy.AtNeutralXY, JoystickPull := joy.AxisCmdY.DirectionPositive, JoystickPush := joy.AxisCmdY.DirectionNegative, BtnValidation := bench.Operator.JoyBtnRaw);
IF bench.Operator.JoyBtnRaw AND NOT previousButton THEN buttonEdges := buttonEdges + 1; END_IF; previousButton := bench.Operator.JoyBtnRaw;
ADVANCE_TIME(10000000);
bench(RawPosM1 := raw1, RawPosM2 := raw2);
joy(RawX := bench.Operator.JoyXRaw_ANA1, RawY := bench.Operator.JoyYRaw_ANA2, RawButton := bench.Operator.JoyBtnRaw, Cfg := cfg, NeutralXMem := nx, NeutralYMem := ny);
home(DeadmanArmed := joy.DeadmanArmed, JoystickDeflected := NOT joy.AtNeutralXY, JoystickPull := joy.AxisCmdY.DirectionPositive, JoystickPush := joy.AxisCmdY.DirectionNegative, BtnValidation := bench.Operator.JoyBtnRaw);
IF bench.Operator.JoyBtnRaw AND NOT previousButton THEN buttonEdges := buttonEdges + 1; END_IF; previousButton := bench.Operator.JoyBtnRaw;
ADVANCE_TIME(10000000);
bench(RawPosM1 := raw1, RawPosM2 := raw2);
joy(RawX := bench.Operator.JoyXRaw_ANA1, RawY := bench.Operator.JoyYRaw_ANA2, RawButton := bench.Operator.JoyBtnRaw, Cfg := cfg, NeutralXMem := nx, NeutralYMem := ny);
home(DeadmanArmed := joy.DeadmanArmed, JoystickDeflected := NOT joy.AtNeutralXY, JoystickPull := joy.AxisCmdY.DirectionPositive, JoystickPush := joy.AxisCmdY.DirectionNegative, BtnValidation := bench.Operator.JoyBtnRaw);
IF bench.Operator.JoyBtnRaw AND NOT previousButton THEN buttonEdges := buttonEdges + 1; END_IF; previousButton := bench.Operator.JoyBtnRaw;
ADVANCE_TIME(10000000);
bench(RawPosM1 := raw1, RawPosM2 := raw2);
joy(RawX := bench.Operator.JoyXRaw_ANA1, RawY := bench.Operator.JoyYRaw_ANA2, RawButton := bench.Operator.JoyBtnRaw, Cfg := cfg, NeutralXMem := nx, NeutralYMem := ny);
home(DeadmanArmed := joy.DeadmanArmed, JoystickDeflected := NOT joy.AtNeutralXY, JoystickPull := joy.AxisCmdY.DirectionPositive, JoystickPush := joy.AxisCmdY.DirectionNegative, BtnValidation := bench.Operator.JoyBtnRaw);
IF bench.Operator.JoyBtnRaw AND NOT previousButton THEN buttonEdges := buttonEdges + 1; END_IF; previousButton := bench.Operator.JoyBtnRaw;
ADVANCE_TIME(10000000);
bench(RawPosM1 := raw1, RawPosM2 := raw2);
joy(RawX := bench.Operator.JoyXRaw_ANA1, RawY := bench.Operator.JoyYRaw_ANA2, RawButton := bench.Operator.JoyBtnRaw, Cfg := cfg, NeutralXMem := nx, NeutralYMem := ny);
home(DeadmanArmed := joy.DeadmanArmed, JoystickDeflected := NOT joy.AtNeutralXY, JoystickPull := joy.AxisCmdY.DirectionPositive, JoystickPush := joy.AxisCmdY.DirectionNegative, BtnValidation := bench.Operator.JoyBtnRaw);
IF bench.Operator.JoyBtnRaw AND NOT previousButton THEN buttonEdges := buttonEdges + 1; END_IF; previousButton := bench.Operator.JoyBtnRaw;
ADVANCE_TIME(10000000);
bench(RawPosM1 := raw1, RawPosM2 := raw2);
joy(RawX := bench.Operator.JoyXRaw_ANA1, RawY := bench.Operator.JoyYRaw_ANA2, RawButton := bench.Operator.JoyBtnRaw, Cfg := cfg, NeutralXMem := nx, NeutralYMem := ny);
home(DeadmanArmed := joy.DeadmanArmed, JoystickDeflected := NOT joy.AtNeutralXY, JoystickPull := joy.AxisCmdY.DirectionPositive, JoystickPush := joy.AxisCmdY.DirectionNegative, BtnValidation := bench.Operator.JoyBtnRaw);
IF bench.Operator.JoyBtnRaw AND NOT previousButton THEN buttonEdges := buttonEdges + 1; END_IF; previousButton := bench.Operator.JoyBtnRaw;
ADVANCE_TIME(10000000);
bench(RawPosM1 := raw1, RawPosM2 := raw2);
joy(RawX := bench.Operator.JoyXRaw_ANA1, RawY := bench.Operator.JoyYRaw_ANA2, RawButton := bench.Operator.JoyBtnRaw, Cfg := cfg, NeutralXMem := nx, NeutralYMem := ny);
home(DeadmanArmed := joy.DeadmanArmed, JoystickDeflected := NOT joy.AtNeutralXY, JoystickPull := joy.AxisCmdY.DirectionPositive, JoystickPush := joy.AxisCmdY.DirectionNegative, BtnValidation := bench.Operator.JoyBtnRaw);
IF bench.Operator.JoyBtnRaw AND NOT previousButton THEN buttonEdges := buttonEdges + 1; END_IF; previousButton := bench.Operator.JoyBtnRaw;
ADVANCE_TIME(10000000);
bench(RawPosM1 := raw1, RawPosM2 := raw2);
joy(RawX := bench.Operator.JoyXRaw_ANA1, RawY := bench.Operator.JoyYRaw_ANA2, RawButton := bench.Operator.JoyBtnRaw, Cfg := cfg, NeutralXMem := nx, NeutralYMem := ny);
home(DeadmanArmed := joy.DeadmanArmed, JoystickDeflected := NOT joy.AtNeutralXY, JoystickPull := joy.AxisCmdY.DirectionPositive, JoystickPush := joy.AxisCmdY.DirectionNegative, BtnValidation := bench.Operator.JoyBtnRaw);
IF bench.Operator.JoyBtnRaw AND NOT previousButton THEN buttonEdges := buttonEdges + 1; END_IF; previousButton := bench.Operator.JoyBtnRaw;
ADVANCE_TIME(10000000);
bench(RawPosM1 := raw1, RawPosM2 := raw2);
joy(RawX := bench.Operator.JoyXRaw_ANA1, RawY := bench.Operator.JoyYRaw_ANA2, RawButton := bench.Operator.JoyBtnRaw, Cfg := cfg, NeutralXMem := nx, NeutralYMem := ny);
home(DeadmanArmed := joy.DeadmanArmed, JoystickDeflected := NOT joy.AtNeutralXY, JoystickPull := joy.AxisCmdY.DirectionPositive, JoystickPush := joy.AxisCmdY.DirectionNegative, BtnValidation := bench.Operator.JoyBtnRaw);
IF bench.Operator.JoyBtnRaw AND NOT previousButton THEN buttonEdges := buttonEdges + 1; END_IF; previousButton := bench.Operator.JoyBtnRaw;
ADVANCE_TIME(10000000);
bench(RawPosM1 := raw1, RawPosM2 := raw2);
joy(RawX := bench.Operator.JoyXRaw_ANA1, RawY := bench.Operator.JoyYRaw_ANA2, RawButton := bench.Operator.JoyBtnRaw, Cfg := cfg, NeutralXMem := nx, NeutralYMem := ny);
home(DeadmanArmed := joy.DeadmanArmed, JoystickDeflected := NOT joy.AtNeutralXY, JoystickPull := joy.AxisCmdY.DirectionPositive, JoystickPush := joy.AxisCmdY.DirectionNegative, BtnValidation := bench.Operator.JoyBtnRaw);
IF bench.Operator.JoyBtnRaw AND NOT previousButton THEN buttonEdges := buttonEdges + 1; END_IF; previousButton := bench.Operator.JoyBtnRaw;
ADVANCE_TIME(10000000);
bench(RawPosM1 := raw1, RawPosM2 := raw2);
joy(RawX := bench.Operator.JoyXRaw_ANA1, RawY := bench.Operator.JoyYRaw_ANA2, RawButton := bench.Operator.JoyBtnRaw, Cfg := cfg, NeutralXMem := nx, NeutralYMem := ny);
home(DeadmanArmed := joy.DeadmanArmed, JoystickDeflected := NOT joy.AtNeutralXY, JoystickPull := joy.AxisCmdY.DirectionPositive, JoystickPush := joy.AxisCmdY.DirectionNegative, BtnValidation := bench.Operator.JoyBtnRaw);
IF bench.Operator.JoyBtnRaw AND NOT previousButton THEN buttonEdges := buttonEdges + 1; END_IF; previousButton := bench.Operator.JoyBtnRaw;
ADVANCE_TIME(10000000);
bench(RawPosM1 := raw1, RawPosM2 := raw2);
joy(RawX := bench.Operator.JoyXRaw_ANA1, RawY := bench.Operator.JoyYRaw_ANA2, RawButton := bench.Operator.JoyBtnRaw, Cfg := cfg, NeutralXMem := nx, NeutralYMem := ny);
home(DeadmanArmed := joy.DeadmanArmed, JoystickDeflected := NOT joy.AtNeutralXY, JoystickPull := joy.AxisCmdY.DirectionPositive, JoystickPush := joy.AxisCmdY.DirectionNegative, BtnValidation := bench.Operator.JoyBtnRaw);
IF bench.Operator.JoyBtnRaw AND NOT previousButton THEN buttonEdges := buttonEdges + 1; END_IF; previousButton := bench.Operator.JoyBtnRaw;
ADVANCE_TIME(10000000);
bench(RawPosM1 := raw1, RawPosM2 := raw2);
joy(RawX := bench.Operator.JoyXRaw_ANA1, RawY := bench.Operator.JoyYRaw_ANA2, RawButton := bench.Operator.JoyBtnRaw, Cfg := cfg, NeutralXMem := nx, NeutralYMem := ny);
home(DeadmanArmed := joy.DeadmanArmed, JoystickDeflected := NOT joy.AtNeutralXY, JoystickPull := joy.AxisCmdY.DirectionPositive, JoystickPush := joy.AxisCmdY.DirectionNegative, BtnValidation := bench.Operator.JoyBtnRaw);
IF bench.Operator.JoyBtnRaw AND NOT previousButton THEN buttonEdges := buttonEdges + 1; END_IF; previousButton := bench.Operator.JoyBtnRaw;
ADVANCE_TIME(10000000);
bench(RawPosM1 := raw1, RawPosM2 := raw2);
joy(RawX := bench.Operator.JoyXRaw_ANA1, RawY := bench.Operator.JoyYRaw_ANA2, RawButton := bench.Operator.JoyBtnRaw, Cfg := cfg, NeutralXMem := nx, NeutralYMem := ny);
home(DeadmanArmed := joy.DeadmanArmed, JoystickDeflected := NOT joy.AtNeutralXY, JoystickPull := joy.AxisCmdY.DirectionPositive, JoystickPush := joy.AxisCmdY.DirectionNegative, BtnValidation := bench.Operator.JoyBtnRaw);
IF bench.Operator.JoyBtnRaw AND NOT previousButton THEN buttonEdges := buttonEdges + 1; END_IF; previousButton := bench.Operator.JoyBtnRaw;
ADVANCE_TIME(10000000);
bench(RawPosM1 := raw1, RawPosM2 := raw2);
joy(RawX := bench.Operator.JoyXRaw_ANA1, RawY := bench.Operator.JoyYRaw_ANA2, RawButton := bench.Operator.JoyBtnRaw, Cfg := cfg, NeutralXMem := nx, NeutralYMem := ny);
home(DeadmanArmed := joy.DeadmanArmed, JoystickDeflected := NOT joy.AtNeutralXY, JoystickPull := joy.AxisCmdY.DirectionPositive, JoystickPush := joy.AxisCmdY.DirectionNegative, BtnValidation := bench.Operator.JoyBtnRaw);
IF bench.Operator.JoyBtnRaw AND NOT previousButton THEN buttonEdges := buttonEdges + 1; END_IF; previousButton := bench.Operator.JoyBtnRaw;
ADVANCE_TIME(10000000);
bench(RawPosM1 := raw1, RawPosM2 := raw2);
joy(RawX := bench.Operator.JoyXRaw_ANA1, RawY := bench.Operator.JoyYRaw_ANA2, RawButton := bench.Operator.JoyBtnRaw, Cfg := cfg, NeutralXMem := nx, NeutralYMem := ny);
home(DeadmanArmed := joy.DeadmanArmed, JoystickDeflected := NOT joy.AtNeutralXY, JoystickPull := joy.AxisCmdY.DirectionPositive, JoystickPush := joy.AxisCmdY.DirectionNegative, BtnValidation := bench.Operator.JoyBtnRaw);
IF bench.Operator.JoyBtnRaw AND NOT previousButton THEN buttonEdges := buttonEdges + 1; END_IF; previousButton := bench.Operator.JoyBtnRaw;
ADVANCE_TIME(10000000);
bench(RawPosM1 := raw1, RawPosM2 := raw2);
joy(RawX := bench.Operator.JoyXRaw_ANA1, RawY := bench.Operator.JoyYRaw_ANA2, RawButton := bench.Operator.JoyBtnRaw, Cfg := cfg, NeutralXMem := nx, NeutralYMem := ny);
home(DeadmanArmed := joy.DeadmanArmed, JoystickDeflected := NOT joy.AtNeutralXY, JoystickPull := joy.AxisCmdY.DirectionPositive, JoystickPush := joy.AxisCmdY.DirectionNegative, BtnValidation := bench.Operator.JoyBtnRaw);
IF bench.Operator.JoyBtnRaw AND NOT previousButton THEN buttonEdges := buttonEdges + 1; END_IF; previousButton := bench.Operator.JoyBtnRaw;
ADVANCE_TIME(10000000);
bench(RawPosM1 := raw1, RawPosM2 := raw2);
joy(RawX := bench.Operator.JoyXRaw_ANA1, RawY := bench.Operator.JoyYRaw_ANA2, RawButton := bench.Operator.JoyBtnRaw, Cfg := cfg, NeutralXMem := nx, NeutralYMem := ny);
home(DeadmanArmed := joy.DeadmanArmed, JoystickDeflected := NOT joy.AtNeutralXY, JoystickPull := joy.AxisCmdY.DirectionPositive, JoystickPush := joy.AxisCmdY.DirectionNegative, BtnValidation := bench.Operator.JoyBtnRaw);
IF bench.Operator.JoyBtnRaw AND NOT previousButton THEN buttonEdges := buttonEdges + 1; END_IF; previousButton := bench.Operator.JoyBtnRaw;
ADVANCE_TIME(10000000);
bench(RawPosM1 := raw1, RawPosM2 := raw2);
joy(RawX := bench.Operator.JoyXRaw_ANA1, RawY := bench.Operator.JoyYRaw_ANA2, RawButton := bench.Operator.JoyBtnRaw, Cfg := cfg, NeutralXMem := nx, NeutralYMem := ny);
home(DeadmanArmed := joy.DeadmanArmed, JoystickDeflected := NOT joy.AtNeutralXY, JoystickPull := joy.AxisCmdY.DirectionPositive, JoystickPush := joy.AxisCmdY.DirectionNegative, BtnValidation := bench.Operator.JoyBtnRaw);
IF bench.Operator.JoyBtnRaw AND NOT previousButton THEN buttonEdges := buttonEdges + 1; END_IF; previousButton := bench.Operator.JoyBtnRaw;
ADVANCE_TIME(10000000);
bench(RawPosM1 := raw1, RawPosM2 := raw2);
joy(RawX := bench.Operator.JoyXRaw_ANA1, RawY := bench.Operator.JoyYRaw_ANA2, RawButton := bench.Operator.JoyBtnRaw, Cfg := cfg, NeutralXMem := nx, NeutralYMem := ny);
home(DeadmanArmed := joy.DeadmanArmed, JoystickDeflected := NOT joy.AtNeutralXY, JoystickPull := joy.AxisCmdY.DirectionPositive, JoystickPush := joy.AxisCmdY.DirectionNegative, BtnValidation := bench.Operator.JoyBtnRaw);
IF bench.Operator.JoyBtnRaw AND NOT previousButton THEN buttonEdges := buttonEdges + 1; END_IF; previousButton := bench.Operator.JoyBtnRaw;
ADVANCE_TIME(10000000);
bench(RawPosM1 := raw1, RawPosM2 := raw2);
joy(RawX := bench.Operator.JoyXRaw_ANA1, RawY := bench.Operator.JoyYRaw_ANA2, RawButton := bench.Operator.JoyBtnRaw, Cfg := cfg, NeutralXMem := nx, NeutralYMem := ny);
home(DeadmanArmed := joy.DeadmanArmed, JoystickDeflected := NOT joy.AtNeutralXY, JoystickPull := joy.AxisCmdY.DirectionPositive, JoystickPush := joy.AxisCmdY.DirectionNegative, BtnValidation := bench.Operator.JoyBtnRaw);
IF bench.Operator.JoyBtnRaw AND NOT previousButton THEN buttonEdges := buttonEdges + 1; END_IF; previousButton := bench.Operator.JoyBtnRaw;
ADVANCE_TIME(10000000);
bench(RawPosM1 := raw1, RawPosM2 := raw2);
joy(RawX := bench.Operator.JoyXRaw_ANA1, RawY := bench.Operator.JoyYRaw_ANA2, RawButton := bench.Operator.JoyBtnRaw, Cfg := cfg, NeutralXMem := nx, NeutralYMem := ny);
home(DeadmanArmed := joy.DeadmanArmed, JoystickDeflected := NOT joy.AtNeutralXY, JoystickPull := joy.AxisCmdY.DirectionPositive, JoystickPush := joy.AxisCmdY.DirectionNegative, BtnValidation := bench.Operator.JoyBtnRaw);
IF bench.Operator.JoyBtnRaw AND NOT previousButton THEN buttonEdges := buttonEdges + 1; END_IF; previousButton := bench.Operator.JoyBtnRaw;
ADVANCE_TIME(10000000);
bench(RawPosM1 := raw1, RawPosM2 := raw2);
joy(RawX := bench.Operator.JoyXRaw_ANA1, RawY := bench.Operator.JoyYRaw_ANA2, RawButton := bench.Operator.JoyBtnRaw, Cfg := cfg, NeutralXMem := nx, NeutralYMem := ny);
home(DeadmanArmed := joy.DeadmanArmed, JoystickDeflected := NOT joy.AtNeutralXY, JoystickPull := joy.AxisCmdY.DirectionPositive, JoystickPush := joy.AxisCmdY.DirectionNegative, BtnValidation := bench.Operator.JoyBtnRaw);
IF bench.Operator.JoyBtnRaw AND NOT previousButton THEN buttonEdges := buttonEdges + 1; END_IF; previousButton := bench.Operator.JoyBtnRaw;
ADVANCE_TIME(10000000);
bench(RawPosM1 := raw1, RawPosM2 := raw2);
joy(RawX := bench.Operator.JoyXRaw_ANA1, RawY := bench.Operator.JoyYRaw_ANA2, RawButton := bench.Operator.JoyBtnRaw, Cfg := cfg, NeutralXMem := nx, NeutralYMem := ny);
home(DeadmanArmed := joy.DeadmanArmed, JoystickDeflected := NOT joy.AtNeutralXY, JoystickPull := joy.AxisCmdY.DirectionPositive, JoystickPush := joy.AxisCmdY.DirectionNegative, BtnValidation := bench.Operator.JoyBtnRaw);
IF bench.Operator.JoyBtnRaw AND NOT previousButton THEN buttonEdges := buttonEdges + 1; END_IF; previousButton := bench.Operator.JoyBtnRaw;
ADVANCE_TIME(10000000);
bench(RawPosM1 := raw1, RawPosM2 := raw2);
joy(RawX := bench.Operator.JoyXRaw_ANA1, RawY := bench.Operator.JoyYRaw_ANA2, RawButton := bench.Operator.JoyBtnRaw, Cfg := cfg, NeutralXMem := nx, NeutralYMem := ny);
home(DeadmanArmed := joy.DeadmanArmed, JoystickDeflected := NOT joy.AtNeutralXY, JoystickPull := joy.AxisCmdY.DirectionPositive, JoystickPush := joy.AxisCmdY.DirectionNegative, BtnValidation := bench.Operator.JoyBtnRaw);
IF bench.Operator.JoyBtnRaw AND NOT previousButton THEN buttonEdges := buttonEdges + 1; END_IF; previousButton := bench.Operator.JoyBtnRaw;
ADVANCE_TIME(10000000);
bench(RawPosM1 := raw1, RawPosM2 := raw2);
joy(RawX := bench.Operator.JoyXRaw_ANA1, RawY := bench.Operator.JoyYRaw_ANA2, RawButton := bench.Operator.JoyBtnRaw, Cfg := cfg, NeutralXMem := nx, NeutralYMem := ny);
home(DeadmanArmed := joy.DeadmanArmed, JoystickDeflected := NOT joy.AtNeutralXY, JoystickPull := joy.AxisCmdY.DirectionPositive, JoystickPush := joy.AxisCmdY.DirectionNegative, BtnValidation := bench.Operator.JoyBtnRaw);
IF bench.Operator.JoyBtnRaw AND NOT previousButton THEN buttonEdges := buttonEdges + 1; END_IF; previousButton := bench.Operator.JoyBtnRaw;
ADVANCE_TIME(10000000);
bench(RawPosM1 := raw1, RawPosM2 := raw2);
joy(RawX := bench.Operator.JoyXRaw_ANA1, RawY := bench.Operator.JoyYRaw_ANA2, RawButton := bench.Operator.JoyBtnRaw, Cfg := cfg, NeutralXMem := nx, NeutralYMem := ny);
home(DeadmanArmed := joy.DeadmanArmed, JoystickDeflected := NOT joy.AtNeutralXY, JoystickPull := joy.AxisCmdY.DirectionPositive, JoystickPush := joy.AxisCmdY.DirectionNegative, BtnValidation := bench.Operator.JoyBtnRaw);
IF bench.Operator.JoyBtnRaw AND NOT previousButton THEN buttonEdges := buttonEdges + 1; END_IF; previousButton := bench.Operator.JoyBtnRaw;
ADVANCE_TIME(10000000);
bench(RawPosM1 := raw1, RawPosM2 := raw2);
joy(RawX := bench.Operator.JoyXRaw_ANA1, RawY := bench.Operator.JoyYRaw_ANA2, RawButton := bench.Operator.JoyBtnRaw, Cfg := cfg, NeutralXMem := nx, NeutralYMem := ny);
home(DeadmanArmed := joy.DeadmanArmed, JoystickDeflected := NOT joy.AtNeutralXY, JoystickPull := joy.AxisCmdY.DirectionPositive, JoystickPush := joy.AxisCmdY.DirectionNegative, BtnValidation := bench.Operator.JoyBtnRaw);
IF bench.Operator.JoyBtnRaw AND NOT previousButton THEN buttonEdges := buttonEdges + 1; END_IF; previousButton := bench.Operator.JoyBtnRaw;
bench.SimJoystickRawX := 9000; bench.SimJoystickRawButton := TRUE; bench.SimJoystickRight_Fwd_MAINT_Active := FALSE;
ADVANCE_TIME(10000000);
bench(RawPosM1 := raw1, RawPosM2 := raw2);
joy(RawX := bench.Operator.JoyXRaw_ANA1, RawY := bench.Operator.JoyYRaw_ANA2, RawButton := bench.Operator.JoyBtnRaw, Cfg := cfg, NeutralXMem := nx, NeutralYMem := ny);
home(DeadmanArmed := joy.DeadmanArmed, JoystickDeflected := NOT joy.AtNeutralXY, JoystickPull := joy.AxisCmdY.DirectionPositive, JoystickPush := joy.AxisCmdY.DirectionNegative, BtnValidation := bench.Operator.JoyBtnRaw);
IF bench.Operator.JoyBtnRaw AND NOT previousButton THEN buttonEdges := buttonEdges + 1; END_IF; previousButton := bench.Operator.JoyBtnRaw;
ADVANCE_TIME(10000000);
bench(RawPosM1 := raw1, RawPosM2 := raw2);
joy(RawX := bench.Operator.JoyXRaw_ANA1, RawY := bench.Operator.JoyYRaw_ANA2, RawButton := bench.Operator.JoyBtnRaw, Cfg := cfg, NeutralXMem := nx, NeutralYMem := ny);
home(DeadmanArmed := joy.DeadmanArmed, JoystickDeflected := NOT joy.AtNeutralXY, JoystickPull := joy.AxisCmdY.DirectionPositive, JoystickPush := joy.AxisCmdY.DirectionNegative, BtnValidation := bench.Operator.JoyBtnRaw);
IF bench.Operator.JoyBtnRaw AND NOT previousButton THEN buttonEdges := buttonEdges + 1; END_IF; previousButton := bench.Operator.JoyBtnRaw;
ADVANCE_TIME(10000000);
bench(RawPosM1 := raw1, RawPosM2 := raw2);
joy(RawX := bench.Operator.JoyXRaw_ANA1, RawY := bench.Operator.JoyYRaw_ANA2, RawButton := bench.Operator.JoyBtnRaw, Cfg := cfg, NeutralXMem := nx, NeutralYMem := ny);
home(DeadmanArmed := joy.DeadmanArmed, JoystickDeflected := NOT joy.AtNeutralXY, JoystickPull := joy.AxisCmdY.DirectionPositive, JoystickPush := joy.AxisCmdY.DirectionNegative, BtnValidation := bench.Operator.JoyBtnRaw);
IF bench.Operator.JoyBtnRaw AND NOT previousButton THEN buttonEdges := buttonEdges + 1; END_IF; previousButton := bench.Operator.JoyBtnRaw;
ADVANCE_TIME(10000000);
bench(RawPosM1 := raw1, RawPosM2 := raw2);
joy(RawX := bench.Operator.JoyXRaw_ANA1, RawY := bench.Operator.JoyYRaw_ANA2, RawButton := bench.Operator.JoyBtnRaw, Cfg := cfg, NeutralXMem := nx, NeutralYMem := ny);
home(DeadmanArmed := joy.DeadmanArmed, JoystickDeflected := NOT joy.AtNeutralXY, JoystickPull := joy.AxisCmdY.DirectionPositive, JoystickPush := joy.AxisCmdY.DirectionNegative, BtnValidation := bench.Operator.JoyBtnRaw);
IF bench.Operator.JoyBtnRaw AND NOT previousButton THEN buttonEdges := buttonEdges + 1; END_IF; previousButton := bench.Operator.JoyBtnRaw;
ADVANCE_TIME(10000000);
bench(RawPosM1 := raw1, RawPosM2 := raw2);
joy(RawX := bench.Operator.JoyXRaw_ANA1, RawY := bench.Operator.JoyYRaw_ANA2, RawButton := bench.Operator.JoyBtnRaw, Cfg := cfg, NeutralXMem := nx, NeutralYMem := ny);
home(DeadmanArmed := joy.DeadmanArmed, JoystickDeflected := NOT joy.AtNeutralXY, JoystickPull := joy.AxisCmdY.DirectionPositive, JoystickPush := joy.AxisCmdY.DirectionNegative, BtnValidation := bench.Operator.JoyBtnRaw);
IF bench.Operator.JoyBtnRaw AND NOT previousButton THEN buttonEdges := buttonEdges + 1; END_IF; previousButton := bench.Operator.JoyBtnRaw;
ADVANCE_TIME(10000000);
bench(RawPosM1 := raw1, RawPosM2 := raw2);
joy(RawX := bench.Operator.JoyXRaw_ANA1, RawY := bench.Operator.JoyYRaw_ANA2, RawButton := bench.Operator.JoyBtnRaw, Cfg := cfg, NeutralXMem := nx, NeutralYMem := ny);
home(DeadmanArmed := joy.DeadmanArmed, JoystickDeflected := NOT joy.AtNeutralXY, JoystickPull := joy.AxisCmdY.DirectionPositive, JoystickPush := joy.AxisCmdY.DirectionNegative, BtnValidation := bench.Operator.JoyBtnRaw);
IF bench.Operator.JoyBtnRaw AND NOT previousButton THEN buttonEdges := buttonEdges + 1; END_IF; previousButton := bench.Operator.JoyBtnRaw;
ADVANCE_TIME(10000000);
bench(RawPosM1 := raw1, RawPosM2 := raw2);
joy(RawX := bench.Operator.JoyXRaw_ANA1, RawY := bench.Operator.JoyYRaw_ANA2, RawButton := bench.Operator.JoyBtnRaw, Cfg := cfg, NeutralXMem := nx, NeutralYMem := ny);
home(DeadmanArmed := joy.DeadmanArmed, JoystickDeflected := NOT joy.AtNeutralXY, JoystickPull := joy.AxisCmdY.DirectionPositive, JoystickPush := joy.AxisCmdY.DirectionNegative, BtnValidation := bench.Operator.JoyBtnRaw);
IF bench.Operator.JoyBtnRaw AND NOT previousButton THEN buttonEdges := buttonEdges + 1; END_IF; previousButton := bench.Operator.JoyBtnRaw;
ADVANCE_TIME(10000000);
bench(RawPosM1 := raw1, RawPosM2 := raw2);
joy(RawX := bench.Operator.JoyXRaw_ANA1, RawY := bench.Operator.JoyYRaw_ANA2, RawButton := bench.Operator.JoyBtnRaw, Cfg := cfg, NeutralXMem := nx, NeutralYMem := ny);
home(DeadmanArmed := joy.DeadmanArmed, JoystickDeflected := NOT joy.AtNeutralXY, JoystickPull := joy.AxisCmdY.DirectionPositive, JoystickPush := joy.AxisCmdY.DirectionNegative, BtnValidation := bench.Operator.JoyBtnRaw);
IF bench.Operator.JoyBtnRaw AND NOT previousButton THEN buttonEdges := buttonEdges + 1; END_IF; previousButton := bench.Operator.JoyBtnRaw;
ADVANCE_TIME(10000000);
bench(RawPosM1 := raw1, RawPosM2 := raw2);
joy(RawX := bench.Operator.JoyXRaw_ANA1, RawY := bench.Operator.JoyYRaw_ANA2, RawButton := bench.Operator.JoyBtnRaw, Cfg := cfg, NeutralXMem := nx, NeutralYMem := ny);
home(DeadmanArmed := joy.DeadmanArmed, JoystickDeflected := NOT joy.AtNeutralXY, JoystickPull := joy.AxisCmdY.DirectionPositive, JoystickPush := joy.AxisCmdY.DirectionNegative, BtnValidation := bench.Operator.JoyBtnRaw);
IF bench.Operator.JoyBtnRaw AND NOT previousButton THEN buttonEdges := buttonEdges + 1; END_IF; previousButton := bench.Operator.JoyBtnRaw;
ADVANCE_TIME(10000000);
bench(RawPosM1 := raw1, RawPosM2 := raw2);
joy(RawX := bench.Operator.JoyXRaw_ANA1, RawY := bench.Operator.JoyYRaw_ANA2, RawButton := bench.Operator.JoyBtnRaw, Cfg := cfg, NeutralXMem := nx, NeutralYMem := ny);
home(DeadmanArmed := joy.DeadmanArmed, JoystickDeflected := NOT joy.AtNeutralXY, JoystickPull := joy.AxisCmdY.DirectionPositive, JoystickPush := joy.AxisCmdY.DirectionNegative, BtnValidation := bench.Operator.JoyBtnRaw);
IF bench.Operator.JoyBtnRaw AND NOT previousButton THEN buttonEdges := buttonEdges + 1; END_IF; previousButton := bench.Operator.JoyBtnRaw;
ADVANCE_TIME(10000000);
bench(RawPosM1 := raw1, RawPosM2 := raw2);
joy(RawX := bench.Operator.JoyXRaw_ANA1, RawY := bench.Operator.JoyYRaw_ANA2, RawButton := bench.Operator.JoyBtnRaw, Cfg := cfg, NeutralXMem := nx, NeutralYMem := ny);
home(DeadmanArmed := joy.DeadmanArmed, JoystickDeflected := NOT joy.AtNeutralXY, JoystickPull := joy.AxisCmdY.DirectionPositive, JoystickPush := joy.AxisCmdY.DirectionNegative, BtnValidation := bench.Operator.JoyBtnRaw);
IF bench.Operator.JoyBtnRaw AND NOT previousButton THEN buttonEdges := buttonEdges + 1; END_IF; previousButton := bench.Operator.JoyBtnRaw;
ADVANCE_TIME(10000000);
bench(RawPosM1 := raw1, RawPosM2 := raw2);
joy(RawX := bench.Operator.JoyXRaw_ANA1, RawY := bench.Operator.JoyYRaw_ANA2, RawButton := bench.Operator.JoyBtnRaw, Cfg := cfg, NeutralXMem := nx, NeutralYMem := ny);
home(DeadmanArmed := joy.DeadmanArmed, JoystickDeflected := NOT joy.AtNeutralXY, JoystickPull := joy.AxisCmdY.DirectionPositive, JoystickPush := joy.AxisCmdY.DirectionNegative, BtnValidation := bench.Operator.JoyBtnRaw);
IF bench.Operator.JoyBtnRaw AND NOT previousButton THEN buttonEdges := buttonEdges + 1; END_IF; previousButton := bench.Operator.JoyBtnRaw;
ADVANCE_TIME(10000000);
bench(RawPosM1 := raw1, RawPosM2 := raw2);
joy(RawX := bench.Operator.JoyXRaw_ANA1, RawY := bench.Operator.JoyYRaw_ANA2, RawButton := bench.Operator.JoyBtnRaw, Cfg := cfg, NeutralXMem := nx, NeutralYMem := ny);
home(DeadmanArmed := joy.DeadmanArmed, JoystickDeflected := NOT joy.AtNeutralXY, JoystickPull := joy.AxisCmdY.DirectionPositive, JoystickPush := joy.AxisCmdY.DirectionNegative, BtnValidation := bench.Operator.JoyBtnRaw);
IF bench.Operator.JoyBtnRaw AND NOT previousButton THEN buttonEdges := buttonEdges + 1; END_IF; previousButton := bench.Operator.JoyBtnRaw;
ADVANCE_TIME(10000000);
bench(RawPosM1 := raw1, RawPosM2 := raw2);
joy(RawX := bench.Operator.JoyXRaw_ANA1, RawY := bench.Operator.JoyYRaw_ANA2, RawButton := bench.Operator.JoyBtnRaw, Cfg := cfg, NeutralXMem := nx, NeutralYMem := ny);
home(DeadmanArmed := joy.DeadmanArmed, JoystickDeflected := NOT joy.AtNeutralXY, JoystickPull := joy.AxisCmdY.DirectionPositive, JoystickPush := joy.AxisCmdY.DirectionNegative, BtnValidation := bench.Operator.JoyBtnRaw);
IF bench.Operator.JoyBtnRaw AND NOT previousButton THEN buttonEdges := buttonEdges + 1; END_IF; previousButton := bench.Operator.JoyBtnRaw;
ADVANCE_TIME(10000000);
bench(RawPosM1 := raw1, RawPosM2 := raw2);
joy(RawX := bench.Operator.JoyXRaw_ANA1, RawY := bench.Operator.JoyYRaw_ANA2, RawButton := bench.Operator.JoyBtnRaw, Cfg := cfg, NeutralXMem := nx, NeutralYMem := ny);
home(DeadmanArmed := joy.DeadmanArmed, JoystickDeflected := NOT joy.AtNeutralXY, JoystickPull := joy.AxisCmdY.DirectionPositive, JoystickPush := joy.AxisCmdY.DirectionNegative, BtnValidation := bench.Operator.JoyBtnRaw);
IF bench.Operator.JoyBtnRaw AND NOT previousButton THEN buttonEdges := buttonEdges + 1; END_IF; previousButton := bench.Operator.JoyBtnRaw;
ADVANCE_TIME(10000000);
bench(RawPosM1 := raw1, RawPosM2 := raw2);
joy(RawX := bench.Operator.JoyXRaw_ANA1, RawY := bench.Operator.JoyYRaw_ANA2, RawButton := bench.Operator.JoyBtnRaw, Cfg := cfg, NeutralXMem := nx, NeutralYMem := ny);
home(DeadmanArmed := joy.DeadmanArmed, JoystickDeflected := NOT joy.AtNeutralXY, JoystickPull := joy.AxisCmdY.DirectionPositive, JoystickPush := joy.AxisCmdY.DirectionNegative, BtnValidation := bench.Operator.JoyBtnRaw);
IF bench.Operator.JoyBtnRaw AND NOT previousButton THEN buttonEdges := buttonEdges + 1; END_IF; previousButton := bench.Operator.JoyBtnRaw;
ADVANCE_TIME(10000000);
bench(RawPosM1 := raw1, RawPosM2 := raw2);
joy(RawX := bench.Operator.JoyXRaw_ANA1, RawY := bench.Operator.JoyYRaw_ANA2, RawButton := bench.Operator.JoyBtnRaw, Cfg := cfg, NeutralXMem := nx, NeutralYMem := ny);
home(DeadmanArmed := joy.DeadmanArmed, JoystickDeflected := NOT joy.AtNeutralXY, JoystickPull := joy.AxisCmdY.DirectionPositive, JoystickPush := joy.AxisCmdY.DirectionNegative, BtnValidation := bench.Operator.JoyBtnRaw);
IF bench.Operator.JoyBtnRaw AND NOT previousButton THEN buttonEdges := buttonEdges + 1; END_IF; previousButton := bench.Operator.JoyBtnRaw;
ADVANCE_TIME(10000000);
bench(RawPosM1 := raw1, RawPosM2 := raw2);
joy(RawX := bench.Operator.JoyXRaw_ANA1, RawY := bench.Operator.JoyYRaw_ANA2, RawButton := bench.Operator.JoyBtnRaw, Cfg := cfg, NeutralXMem := nx, NeutralYMem := ny);
home(DeadmanArmed := joy.DeadmanArmed, JoystickDeflected := NOT joy.AtNeutralXY, JoystickPull := joy.AxisCmdY.DirectionPositive, JoystickPush := joy.AxisCmdY.DirectionNegative, BtnValidation := bench.Operator.JoyBtnRaw);
IF bench.Operator.JoyBtnRaw AND NOT previousButton THEN buttonEdges := buttonEdges + 1; END_IF; previousButton := bench.Operator.JoyBtnRaw;
ADVANCE_TIME(10000000);
bench(RawPosM1 := raw1, RawPosM2 := raw2);
joy(RawX := bench.Operator.JoyXRaw_ANA1, RawY := bench.Operator.JoyYRaw_ANA2, RawButton := bench.Operator.JoyBtnRaw, Cfg := cfg, NeutralXMem := nx, NeutralYMem := ny);
home(DeadmanArmed := joy.DeadmanArmed, JoystickDeflected := NOT joy.AtNeutralXY, JoystickPull := joy.AxisCmdY.DirectionPositive, JoystickPush := joy.AxisCmdY.DirectionNegative, BtnValidation := bench.Operator.JoyBtnRaw);
IF bench.Operator.JoyBtnRaw AND NOT previousButton THEN buttonEdges := buttonEdges + 1; END_IF; previousButton := bench.Operator.JoyBtnRaw;
ADVANCE_TIME(10000000);
bench(RawPosM1 := raw1, RawPosM2 := raw2);
joy(RawX := bench.Operator.JoyXRaw_ANA1, RawY := bench.Operator.JoyYRaw_ANA2, RawButton := bench.Operator.JoyBtnRaw, Cfg := cfg, NeutralXMem := nx, NeutralYMem := ny);
home(DeadmanArmed := joy.DeadmanArmed, JoystickDeflected := NOT joy.AtNeutralXY, JoystickPull := joy.AxisCmdY.DirectionPositive, JoystickPush := joy.AxisCmdY.DirectionNegative, BtnValidation := bench.Operator.JoyBtnRaw);
IF bench.Operator.JoyBtnRaw AND NOT previousButton THEN buttonEdges := buttonEdges + 1; END_IF; previousButton := bench.Operator.JoyBtnRaw;
ADVANCE_TIME(10000000);
bench(RawPosM1 := raw1, RawPosM2 := raw2);
joy(RawX := bench.Operator.JoyXRaw_ANA1, RawY := bench.Operator.JoyYRaw_ANA2, RawButton := bench.Operator.JoyBtnRaw, Cfg := cfg, NeutralXMem := nx, NeutralYMem := ny);
home(DeadmanArmed := joy.DeadmanArmed, JoystickDeflected := NOT joy.AtNeutralXY, JoystickPull := joy.AxisCmdY.DirectionPositive, JoystickPush := joy.AxisCmdY.DirectionNegative, BtnValidation := bench.Operator.JoyBtnRaw);
IF bench.Operator.JoyBtnRaw AND NOT previousButton THEN buttonEdges := buttonEdges + 1; END_IF; previousButton := bench.Operator.JoyBtnRaw;
ADVANCE_TIME(10000000);
bench(RawPosM1 := raw1, RawPosM2 := raw2);
joy(RawX := bench.Operator.JoyXRaw_ANA1, RawY := bench.Operator.JoyYRaw_ANA2, RawButton := bench.Operator.JoyBtnRaw, Cfg := cfg, NeutralXMem := nx, NeutralYMem := ny);
home(DeadmanArmed := joy.DeadmanArmed, JoystickDeflected := NOT joy.AtNeutralXY, JoystickPull := joy.AxisCmdY.DirectionPositive, JoystickPush := joy.AxisCmdY.DirectionNegative, BtnValidation := bench.Operator.JoyBtnRaw);
IF bench.Operator.JoyBtnRaw AND NOT previousButton THEN buttonEdges := buttonEdges + 1; END_IF; previousButton := bench.Operator.JoyBtnRaw;
ADVANCE_TIME(10000000);
bench(RawPosM1 := raw1, RawPosM2 := raw2);
joy(RawX := bench.Operator.JoyXRaw_ANA1, RawY := bench.Operator.JoyYRaw_ANA2, RawButton := bench.Operator.JoyBtnRaw, Cfg := cfg, NeutralXMem := nx, NeutralYMem := ny);
home(DeadmanArmed := joy.DeadmanArmed, JoystickDeflected := NOT joy.AtNeutralXY, JoystickPull := joy.AxisCmdY.DirectionPositive, JoystickPush := joy.AxisCmdY.DirectionNegative, BtnValidation := bench.Operator.JoyBtnRaw);
IF bench.Operator.JoyBtnRaw AND NOT previousButton THEN buttonEdges := buttonEdges + 1; END_IF; previousButton := bench.Operator.JoyBtnRaw;
ADVANCE_TIME(10000000);
bench(RawPosM1 := raw1, RawPosM2 := raw2);
joy(RawX := bench.Operator.JoyXRaw_ANA1, RawY := bench.Operator.JoyYRaw_ANA2, RawButton := bench.Operator.JoyBtnRaw, Cfg := cfg, NeutralXMem := nx, NeutralYMem := ny);
home(DeadmanArmed := joy.DeadmanArmed, JoystickDeflected := NOT joy.AtNeutralXY, JoystickPull := joy.AxisCmdY.DirectionPositive, JoystickPush := joy.AxisCmdY.DirectionNegative, BtnValidation := bench.Operator.JoyBtnRaw);
IF bench.Operator.JoyBtnRaw AND NOT previousButton THEN buttonEdges := buttonEdges + 1; END_IF; previousButton := bench.Operator.JoyBtnRaw;
ADVANCE_TIME(10000000);
bench(RawPosM1 := raw1, RawPosM2 := raw2);
joy(RawX := bench.Operator.JoyXRaw_ANA1, RawY := bench.Operator.JoyYRaw_ANA2, RawButton := bench.Operator.JoyBtnRaw, Cfg := cfg, NeutralXMem := nx, NeutralYMem := ny);
home(DeadmanArmed := joy.DeadmanArmed, JoystickDeflected := NOT joy.AtNeutralXY, JoystickPull := joy.AxisCmdY.DirectionPositive, JoystickPush := joy.AxisCmdY.DirectionNegative, BtnValidation := bench.Operator.JoyBtnRaw);
IF bench.Operator.JoyBtnRaw AND NOT previousButton THEN buttonEdges := buttonEdges + 1; END_IF; previousButton := bench.Operator.JoyBtnRaw;
ADVANCE_TIME(10000000);
bench(RawPosM1 := raw1, RawPosM2 := raw2);
joy(RawX := bench.Operator.JoyXRaw_ANA1, RawY := bench.Operator.JoyYRaw_ANA2, RawButton := bench.Operator.JoyBtnRaw, Cfg := cfg, NeutralXMem := nx, NeutralYMem := ny);
home(DeadmanArmed := joy.DeadmanArmed, JoystickDeflected := NOT joy.AtNeutralXY, JoystickPull := joy.AxisCmdY.DirectionPositive, JoystickPush := joy.AxisCmdY.DirectionNegative, BtnValidation := bench.Operator.JoyBtnRaw);
IF bench.Operator.JoyBtnRaw AND NOT previousButton THEN buttonEdges := buttonEdges + 1; END_IF; previousButton := bench.Operator.JoyBtnRaw;
ADVANCE_TIME(10000000);
bench(RawPosM1 := raw1, RawPosM2 := raw2);
joy(RawX := bench.Operator.JoyXRaw_ANA1, RawY := bench.Operator.JoyYRaw_ANA2, RawButton := bench.Operator.JoyBtnRaw, Cfg := cfg, NeutralXMem := nx, NeutralYMem := ny);
home(DeadmanArmed := joy.DeadmanArmed, JoystickDeflected := NOT joy.AtNeutralXY, JoystickPull := joy.AxisCmdY.DirectionPositive, JoystickPush := joy.AxisCmdY.DirectionNegative, BtnValidation := bench.Operator.JoyBtnRaw);
IF bench.Operator.JoyBtnRaw AND NOT previousButton THEN buttonEdges := buttonEdges + 1; END_IF; previousButton := bench.Operator.JoyBtnRaw;
ADVANCE_TIME(10000000);
bench(RawPosM1 := raw1, RawPosM2 := raw2);
joy(RawX := bench.Operator.JoyXRaw_ANA1, RawY := bench.Operator.JoyYRaw_ANA2, RawButton := bench.Operator.JoyBtnRaw, Cfg := cfg, NeutralXMem := nx, NeutralYMem := ny);
home(DeadmanArmed := joy.DeadmanArmed, JoystickDeflected := NOT joy.AtNeutralXY, JoystickPull := joy.AxisCmdY.DirectionPositive, JoystickPush := joy.AxisCmdY.DirectionNegative, BtnValidation := bench.Operator.JoyBtnRaw);
IF bench.Operator.JoyBtnRaw AND NOT previousButton THEN buttonEdges := buttonEdges + 1; END_IF; previousButton := bench.Operator.JoyBtnRaw;
ADVANCE_TIME(10000000);
bench(RawPosM1 := raw1, RawPosM2 := raw2);
joy(RawX := bench.Operator.JoyXRaw_ANA1, RawY := bench.Operator.JoyYRaw_ANA2, RawButton := bench.Operator.JoyBtnRaw, Cfg := cfg, NeutralXMem := nx, NeutralYMem := ny);
home(DeadmanArmed := joy.DeadmanArmed, JoystickDeflected := NOT joy.AtNeutralXY, JoystickPull := joy.AxisCmdY.DirectionPositive, JoystickPush := joy.AxisCmdY.DirectionNegative, BtnValidation := bench.Operator.JoyBtnRaw);
IF bench.Operator.JoyBtnRaw AND NOT previousButton THEN buttonEdges := buttonEdges + 1; END_IF; previousButton := bench.Operator.JoyBtnRaw;
ADVANCE_TIME(10000000);
bench(RawPosM1 := raw1, RawPosM2 := raw2);
joy(RawX := bench.Operator.JoyXRaw_ANA1, RawY := bench.Operator.JoyYRaw_ANA2, RawButton := bench.Operator.JoyBtnRaw, Cfg := cfg, NeutralXMem := nx, NeutralYMem := ny);
home(DeadmanArmed := joy.DeadmanArmed, JoystickDeflected := NOT joy.AtNeutralXY, JoystickPull := joy.AxisCmdY.DirectionPositive, JoystickPush := joy.AxisCmdY.DirectionNegative, BtnValidation := bench.Operator.JoyBtnRaw);
IF bench.Operator.JoyBtnRaw AND NOT previousButton THEN buttonEdges := buttonEdges + 1; END_IF; previousButton := bench.Operator.JoyBtnRaw;
ADVANCE_TIME(10000000);
bench(RawPosM1 := raw1, RawPosM2 := raw2);
joy(RawX := bench.Operator.JoyXRaw_ANA1, RawY := bench.Operator.JoyYRaw_ANA2, RawButton := bench.Operator.JoyBtnRaw, Cfg := cfg, NeutralXMem := nx, NeutralYMem := ny);
home(DeadmanArmed := joy.DeadmanArmed, JoystickDeflected := NOT joy.AtNeutralXY, JoystickPull := joy.AxisCmdY.DirectionPositive, JoystickPush := joy.AxisCmdY.DirectionNegative, BtnValidation := bench.Operator.JoyBtnRaw);
IF bench.Operator.JoyBtnRaw AND NOT previousButton THEN buttonEdges := buttonEdges + 1; END_IF; previousButton := bench.Operator.JoyBtnRaw;
ADVANCE_TIME(10000000);
bench(RawPosM1 := raw1, RawPosM2 := raw2);
joy(RawX := bench.Operator.JoyXRaw_ANA1, RawY := bench.Operator.JoyYRaw_ANA2, RawButton := bench.Operator.JoyBtnRaw, Cfg := cfg, NeutralXMem := nx, NeutralYMem := ny);
home(DeadmanArmed := joy.DeadmanArmed, JoystickDeflected := NOT joy.AtNeutralXY, JoystickPull := joy.AxisCmdY.DirectionPositive, JoystickPush := joy.AxisCmdY.DirectionNegative, BtnValidation := bench.Operator.JoyBtnRaw);
IF bench.Operator.JoyBtnRaw AND NOT previousButton THEN buttonEdges := buttonEdges + 1; END_IF; previousButton := bench.Operator.JoyBtnRaw;
ADVANCE_TIME(10000000);
bench(RawPosM1 := raw1, RawPosM2 := raw2);
joy(RawX := bench.Operator.JoyXRaw_ANA1, RawY := bench.Operator.JoyYRaw_ANA2, RawButton := bench.Operator.JoyBtnRaw, Cfg := cfg, NeutralXMem := nx, NeutralYMem := ny);
home(DeadmanArmed := joy.DeadmanArmed, JoystickDeflected := NOT joy.AtNeutralXY, JoystickPull := joy.AxisCmdY.DirectionPositive, JoystickPush := joy.AxisCmdY.DirectionNegative, BtnValidation := bench.Operator.JoyBtnRaw);
IF bench.Operator.JoyBtnRaw AND NOT previousButton THEN buttonEdges := buttonEdges + 1; END_IF; previousButton := bench.Operator.JoyBtnRaw;
ADVANCE_TIME(10000000);
bench(RawPosM1 := raw1, RawPosM2 := raw2);
joy(RawX := bench.Operator.JoyXRaw_ANA1, RawY := bench.Operator.JoyYRaw_ANA2, RawButton := bench.Operator.JoyBtnRaw, Cfg := cfg, NeutralXMem := nx, NeutralYMem := ny);
home(DeadmanArmed := joy.DeadmanArmed, JoystickDeflected := NOT joy.AtNeutralXY, JoystickPull := joy.AxisCmdY.DirectionPositive, JoystickPush := joy.AxisCmdY.DirectionNegative, BtnValidation := bench.Operator.JoyBtnRaw);
IF bench.Operator.JoyBtnRaw AND NOT previousButton THEN buttonEdges := buttonEdges + 1; END_IF; previousButton := bench.Operator.JoyBtnRaw;
ADVANCE_TIME(10000000);
bench(RawPosM1 := raw1, RawPosM2 := raw2);
joy(RawX := bench.Operator.JoyXRaw_ANA1, RawY := bench.Operator.JoyYRaw_ANA2, RawButton := bench.Operator.JoyBtnRaw, Cfg := cfg, NeutralXMem := nx, NeutralYMem := ny);
home(DeadmanArmed := joy.DeadmanArmed, JoystickDeflected := NOT joy.AtNeutralXY, JoystickPull := joy.AxisCmdY.DirectionPositive, JoystickPush := joy.AxisCmdY.DirectionNegative, BtnValidation := bench.Operator.JoyBtnRaw);
IF bench.Operator.JoyBtnRaw AND NOT previousButton THEN buttonEdges := buttonEdges + 1; END_IF; previousButton := bench.Operator.JoyBtnRaw;
ASSERT_EQ(bench.Operator.JoyXRaw_ANA1, 5000, 'Fin retour ne saute pas au manuel non neutre'); ASSERT_FALSE(bench.Operator.JoyBtnRaw, 'Bouton manuel bloque pendant conflit');
bench.SimJoystickRawX := 5000; bench.SimJoystickRawButton := FALSE;
ADVANCE_TIME(10000000);
bench(RawPosM1 := raw1, RawPosM2 := raw2);
joy(RawX := bench.Operator.JoyXRaw_ANA1, RawY := bench.Operator.JoyYRaw_ANA2, RawButton := bench.Operator.JoyBtnRaw, Cfg := cfg, NeutralXMem := nx, NeutralYMem := ny);
home(DeadmanArmed := joy.DeadmanArmed, JoystickDeflected := NOT joy.AtNeutralXY, JoystickPull := joy.AxisCmdY.DirectionPositive, JoystickPush := joy.AxisCmdY.DirectionNegative, BtnValidation := bench.Operator.JoyBtnRaw);
IF bench.Operator.JoyBtnRaw AND NOT previousButton THEN buttonEdges := buttonEdges + 1; END_IF; previousButton := bench.Operator.JoyBtnRaw;
END_TEST

TEST 'TC-T418-INT-006 Repli reel puis reactivation banc tenu'
nx := 5000; ny := 5000; raw1 := 0; raw2 := 0; previousButton := FALSE; buttonEdges := 0;
bench.Enable := TRUE; joy.Enable := TRUE; joy.ArmingPermit := TRUE; diagOk.Operational := TRUE;
joy.BusCanOpenOP := diagOk; joy.JoystickOP := diagOk; home.Enable := TRUE; home.BootReady := TRUE;
home.Mode := E_Mode.MAINT_N1; home.BucketOffsetValid := TRUE; home.WinchesMechanicallyStopped := TRUE;
ADVANCE_TIME(10000000);
bench(RawPosM1 := raw1, RawPosM2 := raw2);
joy(RawX := bench.Operator.JoyXRaw_ANA1, RawY := bench.Operator.JoyYRaw_ANA2, RawButton := bench.Operator.JoyBtnRaw, Cfg := cfg, NeutralXMem := nx, NeutralYMem := ny);
home(DeadmanArmed := joy.DeadmanArmed, JoystickDeflected := NOT joy.AtNeutralXY, JoystickPull := joy.AxisCmdY.DirectionPositive, JoystickPush := joy.AxisCmdY.DirectionNegative, BtnValidation := bench.Operator.JoyBtnRaw);
IF bench.Operator.JoyBtnRaw AND NOT previousButton THEN buttonEdges := buttonEdges + 1; END_IF; previousButton := bench.Operator.JoyBtnRaw;
bench.SimJoystickRight_Fwd_MAINT_Active := TRUE;
ADVANCE_TIME(10000000);
bench(RawPosM1 := raw1, RawPosM2 := raw2);
joy(RawX := bench.Operator.JoyXRaw_ANA1, RawY := bench.Operator.JoyYRaw_ANA2, RawButton := bench.Operator.JoyBtnRaw, Cfg := cfg, NeutralXMem := nx, NeutralYMem := ny);
home(DeadmanArmed := joy.DeadmanArmed, JoystickDeflected := NOT joy.AtNeutralXY, JoystickPull := joy.AxisCmdY.DirectionPositive, JoystickPush := joy.AxisCmdY.DirectionNegative, BtnValidation := bench.Operator.JoyBtnRaw);
IF bench.Operator.JoyBtnRaw AND NOT previousButton THEN buttonEdges := buttonEdges + 1; END_IF; previousButton := bench.Operator.JoyBtnRaw;
ADVANCE_TIME(10000000);
bench(RawPosM1 := raw1, RawPosM2 := raw2);
joy(RawX := bench.Operator.JoyXRaw_ANA1, RawY := bench.Operator.JoyYRaw_ANA2, RawButton := bench.Operator.JoyBtnRaw, Cfg := cfg, NeutralXMem := nx, NeutralYMem := ny);
home(DeadmanArmed := joy.DeadmanArmed, JoystickDeflected := NOT joy.AtNeutralXY, JoystickPull := joy.AxisCmdY.DirectionPositive, JoystickPush := joy.AxisCmdY.DirectionNegative, BtnValidation := bench.Operator.JoyBtnRaw);
IF bench.Operator.JoyBtnRaw AND NOT previousButton THEN buttonEdges := buttonEdges + 1; END_IF; previousButton := bench.Operator.JoyBtnRaw;
ADVANCE_TIME(10000000);
bench(RawPosM1 := raw1, RawPosM2 := raw2);
joy(RawX := bench.Operator.JoyXRaw_ANA1, RawY := bench.Operator.JoyYRaw_ANA2, RawButton := bench.Operator.JoyBtnRaw, Cfg := cfg, NeutralXMem := nx, NeutralYMem := ny);
home(DeadmanArmed := joy.DeadmanArmed, JoystickDeflected := NOT joy.AtNeutralXY, JoystickPull := joy.AxisCmdY.DirectionPositive, JoystickPush := joy.AxisCmdY.DirectionNegative, BtnValidation := bench.Operator.JoyBtnRaw);
IF bench.Operator.JoyBtnRaw AND NOT previousButton THEN buttonEdges := buttonEdges + 1; END_IF; previousButton := bench.Operator.JoyBtnRaw;
ADVANCE_TIME(10000000);
bench(RawPosM1 := raw1, RawPosM2 := raw2);
joy(RawX := bench.Operator.JoyXRaw_ANA1, RawY := bench.Operator.JoyYRaw_ANA2, RawButton := bench.Operator.JoyBtnRaw, Cfg := cfg, NeutralXMem := nx, NeutralYMem := ny);
home(DeadmanArmed := joy.DeadmanArmed, JoystickDeflected := NOT joy.AtNeutralXY, JoystickPull := joy.AxisCmdY.DirectionPositive, JoystickPush := joy.AxisCmdY.DirectionNegative, BtnValidation := bench.Operator.JoyBtnRaw);
IF bench.Operator.JoyBtnRaw AND NOT previousButton THEN buttonEdges := buttonEdges + 1; END_IF; previousButton := bench.Operator.JoyBtnRaw;
ADVANCE_TIME(10000000);
bench(RawPosM1 := raw1, RawPosM2 := raw2);
joy(RawX := bench.Operator.JoyXRaw_ANA1, RawY := bench.Operator.JoyYRaw_ANA2, RawButton := bench.Operator.JoyBtnRaw, Cfg := cfg, NeutralXMem := nx, NeutralYMem := ny);
home(DeadmanArmed := joy.DeadmanArmed, JoystickDeflected := NOT joy.AtNeutralXY, JoystickPull := joy.AxisCmdY.DirectionPositive, JoystickPush := joy.AxisCmdY.DirectionNegative, BtnValidation := bench.Operator.JoyBtnRaw);
IF bench.Operator.JoyBtnRaw AND NOT previousButton THEN buttonEdges := buttonEdges + 1; END_IF; previousButton := bench.Operator.JoyBtnRaw;
ADVANCE_TIME(10000000);
bench(RawPosM1 := raw1, RawPosM2 := raw2);
joy(RawX := bench.Operator.JoyXRaw_ANA1, RawY := bench.Operator.JoyYRaw_ANA2, RawButton := bench.Operator.JoyBtnRaw, Cfg := cfg, NeutralXMem := nx, NeutralYMem := ny);
home(DeadmanArmed := joy.DeadmanArmed, JoystickDeflected := NOT joy.AtNeutralXY, JoystickPull := joy.AxisCmdY.DirectionPositive, JoystickPush := joy.AxisCmdY.DirectionNegative, BtnValidation := bench.Operator.JoyBtnRaw);
IF bench.Operator.JoyBtnRaw AND NOT previousButton THEN buttonEdges := buttonEdges + 1; END_IF; previousButton := bench.Operator.JoyBtnRaw;
ADVANCE_TIME(10000000);
bench(RawPosM1 := raw1, RawPosM2 := raw2);
joy(RawX := bench.Operator.JoyXRaw_ANA1, RawY := bench.Operator.JoyYRaw_ANA2, RawButton := bench.Operator.JoyBtnRaw, Cfg := cfg, NeutralXMem := nx, NeutralYMem := ny);
home(DeadmanArmed := joy.DeadmanArmed, JoystickDeflected := NOT joy.AtNeutralXY, JoystickPull := joy.AxisCmdY.DirectionPositive, JoystickPush := joy.AxisCmdY.DirectionNegative, BtnValidation := bench.Operator.JoyBtnRaw);
IF bench.Operator.JoyBtnRaw AND NOT previousButton THEN buttonEdges := buttonEdges + 1; END_IF; previousButton := bench.Operator.JoyBtnRaw;
ADVANCE_TIME(10000000);
bench(RawPosM1 := raw1, RawPosM2 := raw2);
joy(RawX := bench.Operator.JoyXRaw_ANA1, RawY := bench.Operator.JoyYRaw_ANA2, RawButton := bench.Operator.JoyBtnRaw, Cfg := cfg, NeutralXMem := nx, NeutralYMem := ny);
home(DeadmanArmed := joy.DeadmanArmed, JoystickDeflected := NOT joy.AtNeutralXY, JoystickPull := joy.AxisCmdY.DirectionPositive, JoystickPush := joy.AxisCmdY.DirectionNegative, BtnValidation := bench.Operator.JoyBtnRaw);
IF bench.Operator.JoyBtnRaw AND NOT previousButton THEN buttonEdges := buttonEdges + 1; END_IF; previousButton := bench.Operator.JoyBtnRaw;
ADVANCE_TIME(10000000);
bench(RawPosM1 := raw1, RawPosM2 := raw2);
joy(RawX := bench.Operator.JoyXRaw_ANA1, RawY := bench.Operator.JoyYRaw_ANA2, RawButton := bench.Operator.JoyBtnRaw, Cfg := cfg, NeutralXMem := nx, NeutralYMem := ny);
home(DeadmanArmed := joy.DeadmanArmed, JoystickDeflected := NOT joy.AtNeutralXY, JoystickPull := joy.AxisCmdY.DirectionPositive, JoystickPush := joy.AxisCmdY.DirectionNegative, BtnValidation := bench.Operator.JoyBtnRaw);
IF bench.Operator.JoyBtnRaw AND NOT previousButton THEN buttonEdges := buttonEdges + 1; END_IF; previousButton := bench.Operator.JoyBtnRaw;
ADVANCE_TIME(10000000);
bench(RawPosM1 := raw1, RawPosM2 := raw2);
joy(RawX := bench.Operator.JoyXRaw_ANA1, RawY := bench.Operator.JoyYRaw_ANA2, RawButton := bench.Operator.JoyBtnRaw, Cfg := cfg, NeutralXMem := nx, NeutralYMem := ny);
home(DeadmanArmed := joy.DeadmanArmed, JoystickDeflected := NOT joy.AtNeutralXY, JoystickPull := joy.AxisCmdY.DirectionPositive, JoystickPush := joy.AxisCmdY.DirectionNegative, BtnValidation := bench.Operator.JoyBtnRaw);
IF bench.Operator.JoyBtnRaw AND NOT previousButton THEN buttonEdges := buttonEdges + 1; END_IF; previousButton := bench.Operator.JoyBtnRaw;
ADVANCE_TIME(10000000);
bench(RawPosM1 := raw1, RawPosM2 := raw2);
joy(RawX := bench.Operator.JoyXRaw_ANA1, RawY := bench.Operator.JoyYRaw_ANA2, RawButton := bench.Operator.JoyBtnRaw, Cfg := cfg, NeutralXMem := nx, NeutralYMem := ny);
home(DeadmanArmed := joy.DeadmanArmed, JoystickDeflected := NOT joy.AtNeutralXY, JoystickPull := joy.AxisCmdY.DirectionPositive, JoystickPush := joy.AxisCmdY.DirectionNegative, BtnValidation := bench.Operator.JoyBtnRaw);
IF bench.Operator.JoyBtnRaw AND NOT previousButton THEN buttonEdges := buttonEdges + 1; END_IF; previousButton := bench.Operator.JoyBtnRaw;
ADVANCE_TIME(10000000);
bench(RawPosM1 := raw1, RawPosM2 := raw2);
joy(RawX := bench.Operator.JoyXRaw_ANA1, RawY := bench.Operator.JoyYRaw_ANA2, RawButton := bench.Operator.JoyBtnRaw, Cfg := cfg, NeutralXMem := nx, NeutralYMem := ny);
home(DeadmanArmed := joy.DeadmanArmed, JoystickDeflected := NOT joy.AtNeutralXY, JoystickPull := joy.AxisCmdY.DirectionPositive, JoystickPush := joy.AxisCmdY.DirectionNegative, BtnValidation := bench.Operator.JoyBtnRaw);
IF bench.Operator.JoyBtnRaw AND NOT previousButton THEN buttonEdges := buttonEdges + 1; END_IF; previousButton := bench.Operator.JoyBtnRaw;
ADVANCE_TIME(10000000);
bench(RawPosM1 := raw1, RawPosM2 := raw2);
joy(RawX := bench.Operator.JoyXRaw_ANA1, RawY := bench.Operator.JoyYRaw_ANA2, RawButton := bench.Operator.JoyBtnRaw, Cfg := cfg, NeutralXMem := nx, NeutralYMem := ny);
home(DeadmanArmed := joy.DeadmanArmed, JoystickDeflected := NOT joy.AtNeutralXY, JoystickPull := joy.AxisCmdY.DirectionPositive, JoystickPush := joy.AxisCmdY.DirectionNegative, BtnValidation := bench.Operator.JoyBtnRaw);
IF bench.Operator.JoyBtnRaw AND NOT previousButton THEN buttonEdges := buttonEdges + 1; END_IF; previousButton := bench.Operator.JoyBtnRaw;
ADVANCE_TIME(10000000);
bench(RawPosM1 := raw1, RawPosM2 := raw2);
joy(RawX := bench.Operator.JoyXRaw_ANA1, RawY := bench.Operator.JoyYRaw_ANA2, RawButton := bench.Operator.JoyBtnRaw, Cfg := cfg, NeutralXMem := nx, NeutralYMem := ny);
home(DeadmanArmed := joy.DeadmanArmed, JoystickDeflected := NOT joy.AtNeutralXY, JoystickPull := joy.AxisCmdY.DirectionPositive, JoystickPush := joy.AxisCmdY.DirectionNegative, BtnValidation := bench.Operator.JoyBtnRaw);
IF bench.Operator.JoyBtnRaw AND NOT previousButton THEN buttonEdges := buttonEdges + 1; END_IF; previousButton := bench.Operator.JoyBtnRaw;
ADVANCE_TIME(10000000);
bench(RawPosM1 := raw1, RawPosM2 := raw2);
joy(RawX := bench.Operator.JoyXRaw_ANA1, RawY := bench.Operator.JoyYRaw_ANA2, RawButton := bench.Operator.JoyBtnRaw, Cfg := cfg, NeutralXMem := nx, NeutralYMem := ny);
home(DeadmanArmed := joy.DeadmanArmed, JoystickDeflected := NOT joy.AtNeutralXY, JoystickPull := joy.AxisCmdY.DirectionPositive, JoystickPush := joy.AxisCmdY.DirectionNegative, BtnValidation := bench.Operator.JoyBtnRaw);
IF bench.Operator.JoyBtnRaw AND NOT previousButton THEN buttonEdges := buttonEdges + 1; END_IF; previousButton := bench.Operator.JoyBtnRaw;
ADVANCE_TIME(10000000);
bench(RawPosM1 := raw1, RawPosM2 := raw2);
joy(RawX := bench.Operator.JoyXRaw_ANA1, RawY := bench.Operator.JoyYRaw_ANA2, RawButton := bench.Operator.JoyBtnRaw, Cfg := cfg, NeutralXMem := nx, NeutralYMem := ny);
home(DeadmanArmed := joy.DeadmanArmed, JoystickDeflected := NOT joy.AtNeutralXY, JoystickPull := joy.AxisCmdY.DirectionPositive, JoystickPush := joy.AxisCmdY.DirectionNegative, BtnValidation := bench.Operator.JoyBtnRaw);
IF bench.Operator.JoyBtnRaw AND NOT previousButton THEN buttonEdges := buttonEdges + 1; END_IF; previousButton := bench.Operator.JoyBtnRaw;
ADVANCE_TIME(10000000);
bench(RawPosM1 := raw1, RawPosM2 := raw2);
joy(RawX := bench.Operator.JoyXRaw_ANA1, RawY := bench.Operator.JoyYRaw_ANA2, RawButton := bench.Operator.JoyBtnRaw, Cfg := cfg, NeutralXMem := nx, NeutralYMem := ny);
home(DeadmanArmed := joy.DeadmanArmed, JoystickDeflected := NOT joy.AtNeutralXY, JoystickPull := joy.AxisCmdY.DirectionPositive, JoystickPush := joy.AxisCmdY.DirectionNegative, BtnValidation := bench.Operator.JoyBtnRaw);
IF bench.Operator.JoyBtnRaw AND NOT previousButton THEN buttonEdges := buttonEdges + 1; END_IF; previousButton := bench.Operator.JoyBtnRaw;
ADVANCE_TIME(10000000);
bench(RawPosM1 := raw1, RawPosM2 := raw2);
joy(RawX := bench.Operator.JoyXRaw_ANA1, RawY := bench.Operator.JoyYRaw_ANA2, RawButton := bench.Operator.JoyBtnRaw, Cfg := cfg, NeutralXMem := nx, NeutralYMem := ny);
home(DeadmanArmed := joy.DeadmanArmed, JoystickDeflected := NOT joy.AtNeutralXY, JoystickPull := joy.AxisCmdY.DirectionPositive, JoystickPush := joy.AxisCmdY.DirectionNegative, BtnValidation := bench.Operator.JoyBtnRaw);
IF bench.Operator.JoyBtnRaw AND NOT previousButton THEN buttonEdges := buttonEdges + 1; END_IF; previousButton := bench.Operator.JoyBtnRaw;
ADVANCE_TIME(10000000);
bench(RawPosM1 := raw1, RawPosM2 := raw2);
joy(RawX := bench.Operator.JoyXRaw_ANA1, RawY := bench.Operator.JoyYRaw_ANA2, RawButton := bench.Operator.JoyBtnRaw, Cfg := cfg, NeutralXMem := nx, NeutralYMem := ny);
home(DeadmanArmed := joy.DeadmanArmed, JoystickDeflected := NOT joy.AtNeutralXY, JoystickPull := joy.AxisCmdY.DirectionPositive, JoystickPush := joy.AxisCmdY.DirectionNegative, BtnValidation := bench.Operator.JoyBtnRaw);
IF bench.Operator.JoyBtnRaw AND NOT previousButton THEN buttonEdges := buttonEdges + 1; END_IF; previousButton := bench.Operator.JoyBtnRaw;
ADVANCE_TIME(10000000);
bench(RawPosM1 := raw1, RawPosM2 := raw2);
joy(RawX := bench.Operator.JoyXRaw_ANA1, RawY := bench.Operator.JoyYRaw_ANA2, RawButton := bench.Operator.JoyBtnRaw, Cfg := cfg, NeutralXMem := nx, NeutralYMem := ny);
home(DeadmanArmed := joy.DeadmanArmed, JoystickDeflected := NOT joy.AtNeutralXY, JoystickPull := joy.AxisCmdY.DirectionPositive, JoystickPush := joy.AxisCmdY.DirectionNegative, BtnValidation := bench.Operator.JoyBtnRaw);
IF bench.Operator.JoyBtnRaw AND NOT previousButton THEN buttonEdges := buttonEdges + 1; END_IF; previousButton := bench.Operator.JoyBtnRaw;
ADVANCE_TIME(10000000);
bench(RawPosM1 := raw1, RawPosM2 := raw2);
joy(RawX := bench.Operator.JoyXRaw_ANA1, RawY := bench.Operator.JoyYRaw_ANA2, RawButton := bench.Operator.JoyBtnRaw, Cfg := cfg, NeutralXMem := nx, NeutralYMem := ny);
home(DeadmanArmed := joy.DeadmanArmed, JoystickDeflected := NOT joy.AtNeutralXY, JoystickPull := joy.AxisCmdY.DirectionPositive, JoystickPush := joy.AxisCmdY.DirectionNegative, BtnValidation := bench.Operator.JoyBtnRaw);
IF bench.Operator.JoyBtnRaw AND NOT previousButton THEN buttonEdges := buttonEdges + 1; END_IF; previousButton := bench.Operator.JoyBtnRaw;
ADVANCE_TIME(10000000);
bench(RawPosM1 := raw1, RawPosM2 := raw2);
joy(RawX := bench.Operator.JoyXRaw_ANA1, RawY := bench.Operator.JoyYRaw_ANA2, RawButton := bench.Operator.JoyBtnRaw, Cfg := cfg, NeutralXMem := nx, NeutralYMem := ny);
home(DeadmanArmed := joy.DeadmanArmed, JoystickDeflected := NOT joy.AtNeutralXY, JoystickPull := joy.AxisCmdY.DirectionPositive, JoystickPush := joy.AxisCmdY.DirectionNegative, BtnValidation := bench.Operator.JoyBtnRaw);
IF bench.Operator.JoyBtnRaw AND NOT previousButton THEN buttonEdges := buttonEdges + 1; END_IF; previousButton := bench.Operator.JoyBtnRaw;
ADVANCE_TIME(10000000);
bench(RawPosM1 := raw1, RawPosM2 := raw2);
joy(RawX := bench.Operator.JoyXRaw_ANA1, RawY := bench.Operator.JoyYRaw_ANA2, RawButton := bench.Operator.JoyBtnRaw, Cfg := cfg, NeutralXMem := nx, NeutralYMem := ny);
home(DeadmanArmed := joy.DeadmanArmed, JoystickDeflected := NOT joy.AtNeutralXY, JoystickPull := joy.AxisCmdY.DirectionPositive, JoystickPush := joy.AxisCmdY.DirectionNegative, BtnValidation := bench.Operator.JoyBtnRaw);
IF bench.Operator.JoyBtnRaw AND NOT previousButton THEN buttonEdges := buttonEdges + 1; END_IF; previousButton := bench.Operator.JoyBtnRaw;
ADVANCE_TIME(10000000);
bench(RawPosM1 := raw1, RawPosM2 := raw2);
joy(RawX := bench.Operator.JoyXRaw_ANA1, RawY := bench.Operator.JoyYRaw_ANA2, RawButton := bench.Operator.JoyBtnRaw, Cfg := cfg, NeutralXMem := nx, NeutralYMem := ny);
home(DeadmanArmed := joy.DeadmanArmed, JoystickDeflected := NOT joy.AtNeutralXY, JoystickPull := joy.AxisCmdY.DirectionPositive, JoystickPush := joy.AxisCmdY.DirectionNegative, BtnValidation := bench.Operator.JoyBtnRaw);
IF bench.Operator.JoyBtnRaw AND NOT previousButton THEN buttonEdges := buttonEdges + 1; END_IF; previousButton := bench.Operator.JoyBtnRaw;
ADVANCE_TIME(10000000);
bench(RawPosM1 := raw1, RawPosM2 := raw2);
joy(RawX := bench.Operator.JoyXRaw_ANA1, RawY := bench.Operator.JoyYRaw_ANA2, RawButton := bench.Operator.JoyBtnRaw, Cfg := cfg, NeutralXMem := nx, NeutralYMem := ny);
home(DeadmanArmed := joy.DeadmanArmed, JoystickDeflected := NOT joy.AtNeutralXY, JoystickPull := joy.AxisCmdY.DirectionPositive, JoystickPush := joy.AxisCmdY.DirectionNegative, BtnValidation := bench.Operator.JoyBtnRaw);
IF bench.Operator.JoyBtnRaw AND NOT previousButton THEN buttonEdges := buttonEdges + 1; END_IF; previousButton := bench.Operator.JoyBtnRaw;
ADVANCE_TIME(10000000);
bench(RawPosM1 := raw1, RawPosM2 := raw2);
joy(RawX := bench.Operator.JoyXRaw_ANA1, RawY := bench.Operator.JoyYRaw_ANA2, RawButton := bench.Operator.JoyBtnRaw, Cfg := cfg, NeutralXMem := nx, NeutralYMem := ny);
home(DeadmanArmed := joy.DeadmanArmed, JoystickDeflected := NOT joy.AtNeutralXY, JoystickPull := joy.AxisCmdY.DirectionPositive, JoystickPush := joy.AxisCmdY.DirectionNegative, BtnValidation := bench.Operator.JoyBtnRaw);
IF bench.Operator.JoyBtnRaw AND NOT previousButton THEN buttonEdges := buttonEdges + 1; END_IF; previousButton := bench.Operator.JoyBtnRaw;
ADVANCE_TIME(10000000);
bench(RawPosM1 := raw1, RawPosM2 := raw2);
joy(RawX := bench.Operator.JoyXRaw_ANA1, RawY := bench.Operator.JoyYRaw_ANA2, RawButton := bench.Operator.JoyBtnRaw, Cfg := cfg, NeutralXMem := nx, NeutralYMem := ny);
home(DeadmanArmed := joy.DeadmanArmed, JoystickDeflected := NOT joy.AtNeutralXY, JoystickPull := joy.AxisCmdY.DirectionPositive, JoystickPush := joy.AxisCmdY.DirectionNegative, BtnValidation := bench.Operator.JoyBtnRaw);
IF bench.Operator.JoyBtnRaw AND NOT previousButton THEN buttonEdges := buttonEdges + 1; END_IF; previousButton := bench.Operator.JoyBtnRaw;
ADVANCE_TIME(10000000);
bench(RawPosM1 := raw1, RawPosM2 := raw2);
joy(RawX := bench.Operator.JoyXRaw_ANA1, RawY := bench.Operator.JoyYRaw_ANA2, RawButton := bench.Operator.JoyBtnRaw, Cfg := cfg, NeutralXMem := nx, NeutralYMem := ny);
home(DeadmanArmed := joy.DeadmanArmed, JoystickDeflected := NOT joy.AtNeutralXY, JoystickPull := joy.AxisCmdY.DirectionPositive, JoystickPush := joy.AxisCmdY.DirectionNegative, BtnValidation := bench.Operator.JoyBtnRaw);
IF bench.Operator.JoyBtnRaw AND NOT previousButton THEN buttonEdges := buttonEdges + 1; END_IF; previousButton := bench.Operator.JoyBtnRaw;
ADVANCE_TIME(10000000);
bench(RawPosM1 := raw1, RawPosM2 := raw2);
joy(RawX := bench.Operator.JoyXRaw_ANA1, RawY := bench.Operator.JoyYRaw_ANA2, RawButton := bench.Operator.JoyBtnRaw, Cfg := cfg, NeutralXMem := nx, NeutralYMem := ny);
home(DeadmanArmed := joy.DeadmanArmed, JoystickDeflected := NOT joy.AtNeutralXY, JoystickPull := joy.AxisCmdY.DirectionPositive, JoystickPush := joy.AxisCmdY.DirectionNegative, BtnValidation := bench.Operator.JoyBtnRaw);
IF bench.Operator.JoyBtnRaw AND NOT previousButton THEN buttonEdges := buttonEdges + 1; END_IF; previousButton := bench.Operator.JoyBtnRaw;
ADVANCE_TIME(10000000);
bench(RawPosM1 := raw1, RawPosM2 := raw2);
joy(RawX := bench.Operator.JoyXRaw_ANA1, RawY := bench.Operator.JoyYRaw_ANA2, RawButton := bench.Operator.JoyBtnRaw, Cfg := cfg, NeutralXMem := nx, NeutralYMem := ny);
home(DeadmanArmed := joy.DeadmanArmed, JoystickDeflected := NOT joy.AtNeutralXY, JoystickPull := joy.AxisCmdY.DirectionPositive, JoystickPush := joy.AxisCmdY.DirectionNegative, BtnValidation := bench.Operator.JoyBtnRaw);
IF bench.Operator.JoyBtnRaw AND NOT previousButton THEN buttonEdges := buttonEdges + 1; END_IF; previousButton := bench.Operator.JoyBtnRaw;
ADVANCE_TIME(10000000);
bench(RawPosM1 := raw1, RawPosM2 := raw2);
joy(RawX := bench.Operator.JoyXRaw_ANA1, RawY := bench.Operator.JoyYRaw_ANA2, RawButton := bench.Operator.JoyBtnRaw, Cfg := cfg, NeutralXMem := nx, NeutralYMem := ny);
home(DeadmanArmed := joy.DeadmanArmed, JoystickDeflected := NOT joy.AtNeutralXY, JoystickPull := joy.AxisCmdY.DirectionPositive, JoystickPush := joy.AxisCmdY.DirectionNegative, BtnValidation := bench.Operator.JoyBtnRaw);
IF bench.Operator.JoyBtnRaw AND NOT previousButton THEN buttonEdges := buttonEdges + 1; END_IF; previousButton := bench.Operator.JoyBtnRaw;
ADVANCE_TIME(10000000);
bench(RawPosM1 := raw1, RawPosM2 := raw2);
joy(RawX := bench.Operator.JoyXRaw_ANA1, RawY := bench.Operator.JoyYRaw_ANA2, RawButton := bench.Operator.JoyBtnRaw, Cfg := cfg, NeutralXMem := nx, NeutralYMem := ny);
home(DeadmanArmed := joy.DeadmanArmed, JoystickDeflected := NOT joy.AtNeutralXY, JoystickPull := joy.AxisCmdY.DirectionPositive, JoystickPush := joy.AxisCmdY.DirectionNegative, BtnValidation := bench.Operator.JoyBtnRaw);
IF bench.Operator.JoyBtnRaw AND NOT previousButton THEN buttonEdges := buttonEdges + 1; END_IF; previousButton := bench.Operator.JoyBtnRaw;
ADVANCE_TIME(10000000);
bench(RawPosM1 := raw1, RawPosM2 := raw2);
joy(RawX := bench.Operator.JoyXRaw_ANA1, RawY := bench.Operator.JoyYRaw_ANA2, RawButton := bench.Operator.JoyBtnRaw, Cfg := cfg, NeutralXMem := nx, NeutralYMem := ny);
home(DeadmanArmed := joy.DeadmanArmed, JoystickDeflected := NOT joy.AtNeutralXY, JoystickPull := joy.AxisCmdY.DirectionPositive, JoystickPush := joy.AxisCmdY.DirectionNegative, BtnValidation := bench.Operator.JoyBtnRaw);
IF bench.Operator.JoyBtnRaw AND NOT previousButton THEN buttonEdges := buttonEdges + 1; END_IF; previousButton := bench.Operator.JoyBtnRaw;
ADVANCE_TIME(10000000);
bench(RawPosM1 := raw1, RawPosM2 := raw2);
joy(RawX := bench.Operator.JoyXRaw_ANA1, RawY := bench.Operator.JoyYRaw_ANA2, RawButton := bench.Operator.JoyBtnRaw, Cfg := cfg, NeutralXMem := nx, NeutralYMem := ny);
home(DeadmanArmed := joy.DeadmanArmed, JoystickDeflected := NOT joy.AtNeutralXY, JoystickPull := joy.AxisCmdY.DirectionPositive, JoystickPush := joy.AxisCmdY.DirectionNegative, BtnValidation := bench.Operator.JoyBtnRaw);
IF bench.Operator.JoyBtnRaw AND NOT previousButton THEN buttonEdges := buttonEdges + 1; END_IF; previousButton := bench.Operator.JoyBtnRaw;
ADVANCE_TIME(10000000);
bench(RawPosM1 := raw1, RawPosM2 := raw2);
joy(RawX := bench.Operator.JoyXRaw_ANA1, RawY := bench.Operator.JoyYRaw_ANA2, RawButton := bench.Operator.JoyBtnRaw, Cfg := cfg, NeutralXMem := nx, NeutralYMem := ny);
home(DeadmanArmed := joy.DeadmanArmed, JoystickDeflected := NOT joy.AtNeutralXY, JoystickPull := joy.AxisCmdY.DirectionPositive, JoystickPush := joy.AxisCmdY.DirectionNegative, BtnValidation := bench.Operator.JoyBtnRaw);
IF bench.Operator.JoyBtnRaw AND NOT previousButton THEN buttonEdges := buttonEdges + 1; END_IF; previousButton := bench.Operator.JoyBtnRaw;
ADVANCE_TIME(10000000);
bench(RawPosM1 := raw1, RawPosM2 := raw2);
joy(RawX := bench.Operator.JoyXRaw_ANA1, RawY := bench.Operator.JoyYRaw_ANA2, RawButton := bench.Operator.JoyBtnRaw, Cfg := cfg, NeutralXMem := nx, NeutralYMem := ny);
home(DeadmanArmed := joy.DeadmanArmed, JoystickDeflected := NOT joy.AtNeutralXY, JoystickPull := joy.AxisCmdY.DirectionPositive, JoystickPush := joy.AxisCmdY.DirectionNegative, BtnValidation := bench.Operator.JoyBtnRaw);
IF bench.Operator.JoyBtnRaw AND NOT previousButton THEN buttonEdges := buttonEdges + 1; END_IF; previousButton := bench.Operator.JoyBtnRaw;
ADVANCE_TIME(10000000);
bench(RawPosM1 := raw1, RawPosM2 := raw2);
joy(RawX := bench.Operator.JoyXRaw_ANA1, RawY := bench.Operator.JoyYRaw_ANA2, RawButton := bench.Operator.JoyBtnRaw, Cfg := cfg, NeutralXMem := nx, NeutralYMem := ny);
home(DeadmanArmed := joy.DeadmanArmed, JoystickDeflected := NOT joy.AtNeutralXY, JoystickPull := joy.AxisCmdY.DirectionPositive, JoystickPush := joy.AxisCmdY.DirectionNegative, BtnValidation := bench.Operator.JoyBtnRaw);
IF bench.Operator.JoyBtnRaw AND NOT previousButton THEN buttonEdges := buttonEdges + 1; END_IF; previousButton := bench.Operator.JoyBtnRaw;
ADVANCE_TIME(10000000);
bench(RawPosM1 := raw1, RawPosM2 := raw2);
joy(RawX := bench.Operator.JoyXRaw_ANA1, RawY := bench.Operator.JoyYRaw_ANA2, RawButton := bench.Operator.JoyBtnRaw, Cfg := cfg, NeutralXMem := nx, NeutralYMem := ny);
home(DeadmanArmed := joy.DeadmanArmed, JoystickDeflected := NOT joy.AtNeutralXY, JoystickPull := joy.AxisCmdY.DirectionPositive, JoystickPush := joy.AxisCmdY.DirectionNegative, BtnValidation := bench.Operator.JoyBtnRaw);
IF bench.Operator.JoyBtnRaw AND NOT previousButton THEN buttonEdges := buttonEdges + 1; END_IF; previousButton := bench.Operator.JoyBtnRaw;
ADVANCE_TIME(10000000);
bench(RawPosM1 := raw1, RawPosM2 := raw2);
joy(RawX := bench.Operator.JoyXRaw_ANA1, RawY := bench.Operator.JoyYRaw_ANA2, RawButton := bench.Operator.JoyBtnRaw, Cfg := cfg, NeutralXMem := nx, NeutralYMem := ny);
home(DeadmanArmed := joy.DeadmanArmed, JoystickDeflected := NOT joy.AtNeutralXY, JoystickPull := joy.AxisCmdY.DirectionPositive, JoystickPush := joy.AxisCmdY.DirectionNegative, BtnValidation := bench.Operator.JoyBtnRaw);
IF bench.Operator.JoyBtnRaw AND NOT previousButton THEN buttonEdges := buttonEdges + 1; END_IF; previousButton := bench.Operator.JoyBtnRaw;
ADVANCE_TIME(10000000);
bench(RawPosM1 := raw1, RawPosM2 := raw2);
joy(RawX := bench.Operator.JoyXRaw_ANA1, RawY := bench.Operator.JoyYRaw_ANA2, RawButton := bench.Operator.JoyBtnRaw, Cfg := cfg, NeutralXMem := nx, NeutralYMem := ny);
home(DeadmanArmed := joy.DeadmanArmed, JoystickDeflected := NOT joy.AtNeutralXY, JoystickPull := joy.AxisCmdY.DirectionPositive, JoystickPush := joy.AxisCmdY.DirectionNegative, BtnValidation := bench.Operator.JoyBtnRaw);
IF bench.Operator.JoyBtnRaw AND NOT previousButton THEN buttonEdges := buttonEdges + 1; END_IF; previousButton := bench.Operator.JoyBtnRaw;
ADVANCE_TIME(10000000);
bench(RawPosM1 := raw1, RawPosM2 := raw2);
joy(RawX := bench.Operator.JoyXRaw_ANA1, RawY := bench.Operator.JoyYRaw_ANA2, RawButton := bench.Operator.JoyBtnRaw, Cfg := cfg, NeutralXMem := nx, NeutralYMem := ny);
home(DeadmanArmed := joy.DeadmanArmed, JoystickDeflected := NOT joy.AtNeutralXY, JoystickPull := joy.AxisCmdY.DirectionPositive, JoystickPush := joy.AxisCmdY.DirectionNegative, BtnValidation := bench.Operator.JoyBtnRaw);
IF bench.Operator.JoyBtnRaw AND NOT previousButton THEN buttonEdges := buttonEdges + 1; END_IF; previousButton := bench.Operator.JoyBtnRaw;
ADVANCE_TIME(10000000);
bench(RawPosM1 := raw1, RawPosM2 := raw2);
joy(RawX := bench.Operator.JoyXRaw_ANA1, RawY := bench.Operator.JoyYRaw_ANA2, RawButton := bench.Operator.JoyBtnRaw, Cfg := cfg, NeutralXMem := nx, NeutralYMem := ny);
home(DeadmanArmed := joy.DeadmanArmed, JoystickDeflected := NOT joy.AtNeutralXY, JoystickPull := joy.AxisCmdY.DirectionPositive, JoystickPush := joy.AxisCmdY.DirectionNegative, BtnValidation := bench.Operator.JoyBtnRaw);
IF bench.Operator.JoyBtnRaw AND NOT previousButton THEN buttonEdges := buttonEdges + 1; END_IF; previousButton := bench.Operator.JoyBtnRaw;
ADVANCE_TIME(10000000);
bench(RawPosM1 := raw1, RawPosM2 := raw2);
joy(RawX := bench.Operator.JoyXRaw_ANA1, RawY := bench.Operator.JoyYRaw_ANA2, RawButton := bench.Operator.JoyBtnRaw, Cfg := cfg, NeutralXMem := nx, NeutralYMem := ny);
home(DeadmanArmed := joy.DeadmanArmed, JoystickDeflected := NOT joy.AtNeutralXY, JoystickPull := joy.AxisCmdY.DirectionPositive, JoystickPush := joy.AxisCmdY.DirectionNegative, BtnValidation := bench.Operator.JoyBtnRaw);
IF bench.Operator.JoyBtnRaw AND NOT previousButton THEN buttonEdges := buttonEdges + 1; END_IF; previousButton := bench.Operator.JoyBtnRaw;
ADVANCE_TIME(10000000);
bench(RawPosM1 := raw1, RawPosM2 := raw2);
joy(RawX := bench.Operator.JoyXRaw_ANA1, RawY := bench.Operator.JoyYRaw_ANA2, RawButton := bench.Operator.JoyBtnRaw, Cfg := cfg, NeutralXMem := nx, NeutralYMem := ny);
home(DeadmanArmed := joy.DeadmanArmed, JoystickDeflected := NOT joy.AtNeutralXY, JoystickPull := joy.AxisCmdY.DirectionPositive, JoystickPush := joy.AxisCmdY.DirectionNegative, BtnValidation := bench.Operator.JoyBtnRaw);
IF bench.Operator.JoyBtnRaw AND NOT previousButton THEN buttonEdges := buttonEdges + 1; END_IF; previousButton := bench.Operator.JoyBtnRaw;
ADVANCE_TIME(10000000);
bench(RawPosM1 := raw1, RawPosM2 := raw2);
joy(RawX := bench.Operator.JoyXRaw_ANA1, RawY := bench.Operator.JoyYRaw_ANA2, RawButton := bench.Operator.JoyBtnRaw, Cfg := cfg, NeutralXMem := nx, NeutralYMem := ny);
home(DeadmanArmed := joy.DeadmanArmed, JoystickDeflected := NOT joy.AtNeutralXY, JoystickPull := joy.AxisCmdY.DirectionPositive, JoystickPush := joy.AxisCmdY.DirectionNegative, BtnValidation := bench.Operator.JoyBtnRaw);
IF bench.Operator.JoyBtnRaw AND NOT previousButton THEN buttonEdges := buttonEdges + 1; END_IF; previousButton := bench.Operator.JoyBtnRaw;
ADVANCE_TIME(10000000);
bench(RawPosM1 := raw1, RawPosM2 := raw2);
joy(RawX := bench.Operator.JoyXRaw_ANA1, RawY := bench.Operator.JoyYRaw_ANA2, RawButton := bench.Operator.JoyBtnRaw, Cfg := cfg, NeutralXMem := nx, NeutralYMem := ny);
home(DeadmanArmed := joy.DeadmanArmed, JoystickDeflected := NOT joy.AtNeutralXY, JoystickPull := joy.AxisCmdY.DirectionPositive, JoystickPush := joy.AxisCmdY.DirectionNegative, BtnValidation := bench.Operator.JoyBtnRaw);
IF bench.Operator.JoyBtnRaw AND NOT previousButton THEN buttonEdges := buttonEdges + 1; END_IF; previousButton := bench.Operator.JoyBtnRaw;
ADVANCE_TIME(10000000);
bench(RawPosM1 := raw1, RawPosM2 := raw2);
joy(RawX := bench.Operator.JoyXRaw_ANA1, RawY := bench.Operator.JoyYRaw_ANA2, RawButton := bench.Operator.JoyBtnRaw, Cfg := cfg, NeutralXMem := nx, NeutralYMem := ny);
home(DeadmanArmed := joy.DeadmanArmed, JoystickDeflected := NOT joy.AtNeutralXY, JoystickPull := joy.AxisCmdY.DirectionPositive, JoystickPush := joy.AxisCmdY.DirectionNegative, BtnValidation := bench.Operator.JoyBtnRaw);
IF bench.Operator.JoyBtnRaw AND NOT previousButton THEN buttonEdges := buttonEdges + 1; END_IF; previousButton := bench.Operator.JoyBtnRaw;
ADVANCE_TIME(10000000);
bench(RawPosM1 := raw1, RawPosM2 := raw2);
joy(RawX := bench.Operator.JoyXRaw_ANA1, RawY := bench.Operator.JoyYRaw_ANA2, RawButton := bench.Operator.JoyBtnRaw, Cfg := cfg, NeutralXMem := nx, NeutralYMem := ny);
home(DeadmanArmed := joy.DeadmanArmed, JoystickDeflected := NOT joy.AtNeutralXY, JoystickPull := joy.AxisCmdY.DirectionPositive, JoystickPush := joy.AxisCmdY.DirectionNegative, BtnValidation := bench.Operator.JoyBtnRaw);
IF bench.Operator.JoyBtnRaw AND NOT previousButton THEN buttonEdges := buttonEdges + 1; END_IF; previousButton := bench.Operator.JoyBtnRaw;
ADVANCE_TIME(10000000);
bench(RawPosM1 := raw1, RawPosM2 := raw2);
joy(RawX := bench.Operator.JoyXRaw_ANA1, RawY := bench.Operator.JoyYRaw_ANA2, RawButton := bench.Operator.JoyBtnRaw, Cfg := cfg, NeutralXMem := nx, NeutralYMem := ny);
home(DeadmanArmed := joy.DeadmanArmed, JoystickDeflected := NOT joy.AtNeutralXY, JoystickPull := joy.AxisCmdY.DirectionPositive, JoystickPush := joy.AxisCmdY.DirectionNegative, BtnValidation := bench.Operator.JoyBtnRaw);
IF bench.Operator.JoyBtnRaw AND NOT previousButton THEN buttonEdges := buttonEdges + 1; END_IF; previousButton := bench.Operator.JoyBtnRaw;
ADVANCE_TIME(10000000);
bench(RawPosM1 := raw1, RawPosM2 := raw2);
joy(RawX := bench.Operator.JoyXRaw_ANA1, RawY := bench.Operator.JoyYRaw_ANA2, RawButton := bench.Operator.JoyBtnRaw, Cfg := cfg, NeutralXMem := nx, NeutralYMem := ny);
home(DeadmanArmed := joy.DeadmanArmed, JoystickDeflected := NOT joy.AtNeutralXY, JoystickPull := joy.AxisCmdY.DirectionPositive, JoystickPush := joy.AxisCmdY.DirectionNegative, BtnValidation := bench.Operator.JoyBtnRaw);
IF bench.Operator.JoyBtnRaw AND NOT previousButton THEN buttonEdges := buttonEdges + 1; END_IF; previousButton := bench.Operator.JoyBtnRaw;
ADVANCE_TIME(10000000);
bench(RawPosM1 := raw1, RawPosM2 := raw2);
joy(RawX := bench.Operator.JoyXRaw_ANA1, RawY := bench.Operator.JoyYRaw_ANA2, RawButton := bench.Operator.JoyBtnRaw, Cfg := cfg, NeutralXMem := nx, NeutralYMem := ny);
home(DeadmanArmed := joy.DeadmanArmed, JoystickDeflected := NOT joy.AtNeutralXY, JoystickPull := joy.AxisCmdY.DirectionPositive, JoystickPush := joy.AxisCmdY.DirectionNegative, BtnValidation := bench.Operator.JoyBtnRaw);
IF bench.Operator.JoyBtnRaw AND NOT previousButton THEN buttonEdges := buttonEdges + 1; END_IF; previousButton := bench.Operator.JoyBtnRaw;
ADVANCE_TIME(10000000);
bench(RawPosM1 := raw1, RawPosM2 := raw2);
joy(RawX := bench.Operator.JoyXRaw_ANA1, RawY := bench.Operator.JoyYRaw_ANA2, RawButton := bench.Operator.JoyBtnRaw, Cfg := cfg, NeutralXMem := nx, NeutralYMem := ny);
home(DeadmanArmed := joy.DeadmanArmed, JoystickDeflected := NOT joy.AtNeutralXY, JoystickPull := joy.AxisCmdY.DirectionPositive, JoystickPush := joy.AxisCmdY.DirectionNegative, BtnValidation := bench.Operator.JoyBtnRaw);
IF bench.Operator.JoyBtnRaw AND NOT previousButton THEN buttonEdges := buttonEdges + 1; END_IF; previousButton := bench.Operator.JoyBtnRaw;
ADVANCE_TIME(10000000);
bench(RawPosM1 := raw1, RawPosM2 := raw2);
joy(RawX := bench.Operator.JoyXRaw_ANA1, RawY := bench.Operator.JoyYRaw_ANA2, RawButton := bench.Operator.JoyBtnRaw, Cfg := cfg, NeutralXMem := nx, NeutralYMem := ny);
home(DeadmanArmed := joy.DeadmanArmed, JoystickDeflected := NOT joy.AtNeutralXY, JoystickPull := joy.AxisCmdY.DirectionPositive, JoystickPush := joy.AxisCmdY.DirectionNegative, BtnValidation := bench.Operator.JoyBtnRaw);
IF bench.Operator.JoyBtnRaw AND NOT previousButton THEN buttonEdges := buttonEdges + 1; END_IF; previousButton := bench.Operator.JoyBtnRaw;
ADVANCE_TIME(10000000);
bench(RawPosM1 := raw1, RawPosM2 := raw2);
joy(RawX := bench.Operator.JoyXRaw_ANA1, RawY := bench.Operator.JoyYRaw_ANA2, RawButton := bench.Operator.JoyBtnRaw, Cfg := cfg, NeutralXMem := nx, NeutralYMem := ny);
home(DeadmanArmed := joy.DeadmanArmed, JoystickDeflected := NOT joy.AtNeutralXY, JoystickPull := joy.AxisCmdY.DirectionPositive, JoystickPush := joy.AxisCmdY.DirectionNegative, BtnValidation := bench.Operator.JoyBtnRaw);
IF bench.Operator.JoyBtnRaw AND NOT previousButton THEN buttonEdges := buttonEdges + 1; END_IF; previousButton := bench.Operator.JoyBtnRaw;
ADVANCE_TIME(10000000);
bench(RawPosM1 := raw1, RawPosM2 := raw2);
joy(RawX := bench.Operator.JoyXRaw_ANA1, RawY := bench.Operator.JoyYRaw_ANA2, RawButton := bench.Operator.JoyBtnRaw, Cfg := cfg, NeutralXMem := nx, NeutralYMem := ny);
home(DeadmanArmed := joy.DeadmanArmed, JoystickDeflected := NOT joy.AtNeutralXY, JoystickPull := joy.AxisCmdY.DirectionPositive, JoystickPush := joy.AxisCmdY.DirectionNegative, BtnValidation := bench.Operator.JoyBtnRaw);
IF bench.Operator.JoyBtnRaw AND NOT previousButton THEN buttonEdges := buttonEdges + 1; END_IF; previousButton := bench.Operator.JoyBtnRaw;
ADVANCE_TIME(10000000);
bench(RawPosM1 := raw1, RawPosM2 := raw2);
joy(RawX := bench.Operator.JoyXRaw_ANA1, RawY := bench.Operator.JoyYRaw_ANA2, RawButton := bench.Operator.JoyBtnRaw, Cfg := cfg, NeutralXMem := nx, NeutralYMem := ny);
home(DeadmanArmed := joy.DeadmanArmed, JoystickDeflected := NOT joy.AtNeutralXY, JoystickPull := joy.AxisCmdY.DirectionPositive, JoystickPush := joy.AxisCmdY.DirectionNegative, BtnValidation := bench.Operator.JoyBtnRaw);
IF bench.Operator.JoyBtnRaw AND NOT previousButton THEN buttonEdges := buttonEdges + 1; END_IF; previousButton := bench.Operator.JoyBtnRaw;
ADVANCE_TIME(10000000);
bench(RawPosM1 := raw1, RawPosM2 := raw2);
joy(RawX := bench.Operator.JoyXRaw_ANA1, RawY := bench.Operator.JoyYRaw_ANA2, RawButton := bench.Operator.JoyBtnRaw, Cfg := cfg, NeutralXMem := nx, NeutralYMem := ny);
home(DeadmanArmed := joy.DeadmanArmed, JoystickDeflected := NOT joy.AtNeutralXY, JoystickPull := joy.AxisCmdY.DirectionPositive, JoystickPush := joy.AxisCmdY.DirectionNegative, BtnValidation := bench.Operator.JoyBtnRaw);
IF bench.Operator.JoyBtnRaw AND NOT previousButton THEN buttonEdges := buttonEdges + 1; END_IF; previousButton := bench.Operator.JoyBtnRaw;
ADVANCE_TIME(10000000);
bench(RawPosM1 := raw1, RawPosM2 := raw2);
joy(RawX := bench.Operator.JoyXRaw_ANA1, RawY := bench.Operator.JoyYRaw_ANA2, RawButton := bench.Operator.JoyBtnRaw, Cfg := cfg, NeutralXMem := nx, NeutralYMem := ny);
home(DeadmanArmed := joy.DeadmanArmed, JoystickDeflected := NOT joy.AtNeutralXY, JoystickPull := joy.AxisCmdY.DirectionPositive, JoystickPush := joy.AxisCmdY.DirectionNegative, BtnValidation := bench.Operator.JoyBtnRaw);
IF bench.Operator.JoyBtnRaw AND NOT previousButton THEN buttonEdges := buttonEdges + 1; END_IF; previousButton := bench.Operator.JoyBtnRaw;
ADVANCE_TIME(10000000);
bench(RawPosM1 := raw1, RawPosM2 := raw2);
joy(RawX := bench.Operator.JoyXRaw_ANA1, RawY := bench.Operator.JoyYRaw_ANA2, RawButton := bench.Operator.JoyBtnRaw, Cfg := cfg, NeutralXMem := nx, NeutralYMem := ny);
home(DeadmanArmed := joy.DeadmanArmed, JoystickDeflected := NOT joy.AtNeutralXY, JoystickPull := joy.AxisCmdY.DirectionPositive, JoystickPush := joy.AxisCmdY.DirectionNegative, BtnValidation := bench.Operator.JoyBtnRaw);
IF bench.Operator.JoyBtnRaw AND NOT previousButton THEN buttonEdges := buttonEdges + 1; END_IF; previousButton := bench.Operator.JoyBtnRaw;
ADVANCE_TIME(10000000);
bench(RawPosM1 := raw1, RawPosM2 := raw2);
joy(RawX := bench.Operator.JoyXRaw_ANA1, RawY := bench.Operator.JoyYRaw_ANA2, RawButton := bench.Operator.JoyBtnRaw, Cfg := cfg, NeutralXMem := nx, NeutralYMem := ny);
home(DeadmanArmed := joy.DeadmanArmed, JoystickDeflected := NOT joy.AtNeutralXY, JoystickPull := joy.AxisCmdY.DirectionPositive, JoystickPush := joy.AxisCmdY.DirectionNegative, BtnValidation := bench.Operator.JoyBtnRaw);
IF bench.Operator.JoyBtnRaw AND NOT previousButton THEN buttonEdges := buttonEdges + 1; END_IF; previousButton := bench.Operator.JoyBtnRaw;
ADVANCE_TIME(10000000);
bench(RawPosM1 := raw1, RawPosM2 := raw2);
joy(RawX := bench.Operator.JoyXRaw_ANA1, RawY := bench.Operator.JoyYRaw_ANA2, RawButton := bench.Operator.JoyBtnRaw, Cfg := cfg, NeutralXMem := nx, NeutralYMem := ny);
home(DeadmanArmed := joy.DeadmanArmed, JoystickDeflected := NOT joy.AtNeutralXY, JoystickPull := joy.AxisCmdY.DirectionPositive, JoystickPush := joy.AxisCmdY.DirectionNegative, BtnValidation := bench.Operator.JoyBtnRaw);
IF bench.Operator.JoyBtnRaw AND NOT previousButton THEN buttonEdges := buttonEdges + 1; END_IF; previousButton := bench.Operator.JoyBtnRaw;
ADVANCE_TIME(10000000);
bench(RawPosM1 := raw1, RawPosM2 := raw2);
joy(RawX := bench.Operator.JoyXRaw_ANA1, RawY := bench.Operator.JoyYRaw_ANA2, RawButton := bench.Operator.JoyBtnRaw, Cfg := cfg, NeutralXMem := nx, NeutralYMem := ny);
home(DeadmanArmed := joy.DeadmanArmed, JoystickDeflected := NOT joy.AtNeutralXY, JoystickPull := joy.AxisCmdY.DirectionPositive, JoystickPush := joy.AxisCmdY.DirectionNegative, BtnValidation := bench.Operator.JoyBtnRaw);
IF bench.Operator.JoyBtnRaw AND NOT previousButton THEN buttonEdges := buttonEdges + 1; END_IF; previousButton := bench.Operator.JoyBtnRaw;
ADVANCE_TIME(10000000);
bench(RawPosM1 := raw1, RawPosM2 := raw2);
joy(RawX := bench.Operator.JoyXRaw_ANA1, RawY := bench.Operator.JoyYRaw_ANA2, RawButton := bench.Operator.JoyBtnRaw, Cfg := cfg, NeutralXMem := nx, NeutralYMem := ny);
home(DeadmanArmed := joy.DeadmanArmed, JoystickDeflected := NOT joy.AtNeutralXY, JoystickPull := joy.AxisCmdY.DirectionPositive, JoystickPush := joy.AxisCmdY.DirectionNegative, BtnValidation := bench.Operator.JoyBtnRaw);
IF bench.Operator.JoyBtnRaw AND NOT previousButton THEN buttonEdges := buttonEdges + 1; END_IF; previousButton := bench.Operator.JoyBtnRaw;
ADVANCE_TIME(10000000);
bench(RawPosM1 := raw1, RawPosM2 := raw2);
joy(RawX := bench.Operator.JoyXRaw_ANA1, RawY := bench.Operator.JoyYRaw_ANA2, RawButton := bench.Operator.JoyBtnRaw, Cfg := cfg, NeutralXMem := nx, NeutralYMem := ny);
home(DeadmanArmed := joy.DeadmanArmed, JoystickDeflected := NOT joy.AtNeutralXY, JoystickPull := joy.AxisCmdY.DirectionPositive, JoystickPush := joy.AxisCmdY.DirectionNegative, BtnValidation := bench.Operator.JoyBtnRaw);
IF bench.Operator.JoyBtnRaw AND NOT previousButton THEN buttonEdges := buttonEdges + 1; END_IF; previousButton := bench.Operator.JoyBtnRaw;
ADVANCE_TIME(10000000);
bench(RawPosM1 := raw1, RawPosM2 := raw2);
joy(RawX := bench.Operator.JoyXRaw_ANA1, RawY := bench.Operator.JoyYRaw_ANA2, RawButton := bench.Operator.JoyBtnRaw, Cfg := cfg, NeutralXMem := nx, NeutralYMem := ny);
home(DeadmanArmed := joy.DeadmanArmed, JoystickDeflected := NOT joy.AtNeutralXY, JoystickPull := joy.AxisCmdY.DirectionPositive, JoystickPush := joy.AxisCmdY.DirectionNegative, BtnValidation := bench.Operator.JoyBtnRaw);
IF bench.Operator.JoyBtnRaw AND NOT previousButton THEN buttonEdges := buttonEdges + 1; END_IF; previousButton := bench.Operator.JoyBtnRaw;
bench.Enable := FALSE; bench.HwReal.Operator.JoyXRaw_ANA1 := 4321; bench.HwReal.Operator.JoyBtnRaw := TRUE;
ADVANCE_TIME(10000000);
bench(RawPosM1 := raw1, RawPosM2 := raw2);
joy(RawX := bench.Operator.JoyXRaw_ANA1, RawY := bench.Operator.JoyYRaw_ANA2, RawButton := bench.Operator.JoyBtnRaw, Cfg := cfg, NeutralXMem := nx, NeutralYMem := ny);
home(DeadmanArmed := joy.DeadmanArmed, JoystickDeflected := NOT joy.AtNeutralXY, JoystickPull := joy.AxisCmdY.DirectionPositive, JoystickPush := joy.AxisCmdY.DirectionNegative, BtnValidation := bench.Operator.JoyBtnRaw);
IF bench.Operator.JoyBtnRaw AND NOT previousButton THEN buttonEdges := buttonEdges + 1; END_IF; previousButton := bench.Operator.JoyBtnRaw;
ASSERT_EQ(bench.Operator.JoyXRaw_ANA1, 4321, 'Repli image reelle conserve'); ASSERT_TRUE(bench.Operator.JoyBtnRaw, 'Bouton reel conserve hors banc');
bench.Enable := TRUE;
ADVANCE_TIME(10000000);
bench(RawPosM1 := raw1, RawPosM2 := raw2);
joy(RawX := bench.Operator.JoyXRaw_ANA1, RawY := bench.Operator.JoyYRaw_ANA2, RawButton := bench.Operator.JoyBtnRaw, Cfg := cfg, NeutralXMem := nx, NeutralYMem := ny);
home(DeadmanArmed := joy.DeadmanArmed, JoystickDeflected := NOT joy.AtNeutralXY, JoystickPull := joy.AxisCmdY.DirectionPositive, JoystickPush := joy.AxisCmdY.DirectionNegative, BtnValidation := bench.Operator.JoyBtnRaw);
IF bench.Operator.JoyBtnRaw AND NOT previousButton THEN buttonEdges := buttonEdges + 1; END_IF; previousButton := bench.Operator.JoyBtnRaw;
ASSERT_EQ(bench.Operator.JoyXRaw_ANA1, 5000, 'Pas de reprise apres OFF ON'); ASSERT_FALSE(bench.Operator.JoyBtnRaw, 'Bouton tenu ignore');
ADVANCE_TIME(10000000);
bench(RawPosM1 := raw1, RawPosM2 := raw2);
joy(RawX := bench.Operator.JoyXRaw_ANA1, RawY := bench.Operator.JoyYRaw_ANA2, RawButton := bench.Operator.JoyBtnRaw, Cfg := cfg, NeutralXMem := nx, NeutralYMem := ny);
home(DeadmanArmed := joy.DeadmanArmed, JoystickDeflected := NOT joy.AtNeutralXY, JoystickPull := joy.AxisCmdY.DirectionPositive, JoystickPush := joy.AxisCmdY.DirectionNegative, BtnValidation := bench.Operator.JoyBtnRaw);
IF bench.Operator.JoyBtnRaw AND NOT previousButton THEN buttonEdges := buttonEdges + 1; END_IF; previousButton := bench.Operator.JoyBtnRaw;
ASSERT_EQ(bench.Operator.JoyXRaw_ANA1, 5000, 'Pas de reprise apres OFF ON'); ASSERT_FALSE(bench.Operator.JoyBtnRaw, 'Bouton tenu ignore');
ADVANCE_TIME(10000000);
bench(RawPosM1 := raw1, RawPosM2 := raw2);
joy(RawX := bench.Operator.JoyXRaw_ANA1, RawY := bench.Operator.JoyYRaw_ANA2, RawButton := bench.Operator.JoyBtnRaw, Cfg := cfg, NeutralXMem := nx, NeutralYMem := ny);
home(DeadmanArmed := joy.DeadmanArmed, JoystickDeflected := NOT joy.AtNeutralXY, JoystickPull := joy.AxisCmdY.DirectionPositive, JoystickPush := joy.AxisCmdY.DirectionNegative, BtnValidation := bench.Operator.JoyBtnRaw);
IF bench.Operator.JoyBtnRaw AND NOT previousButton THEN buttonEdges := buttonEdges + 1; END_IF; previousButton := bench.Operator.JoyBtnRaw;
ASSERT_EQ(bench.Operator.JoyXRaw_ANA1, 5000, 'Pas de reprise apres OFF ON'); ASSERT_FALSE(bench.Operator.JoyBtnRaw, 'Bouton tenu ignore');
ADVANCE_TIME(10000000);
bench(RawPosM1 := raw1, RawPosM2 := raw2);
joy(RawX := bench.Operator.JoyXRaw_ANA1, RawY := bench.Operator.JoyYRaw_ANA2, RawButton := bench.Operator.JoyBtnRaw, Cfg := cfg, NeutralXMem := nx, NeutralYMem := ny);
home(DeadmanArmed := joy.DeadmanArmed, JoystickDeflected := NOT joy.AtNeutralXY, JoystickPull := joy.AxisCmdY.DirectionPositive, JoystickPush := joy.AxisCmdY.DirectionNegative, BtnValidation := bench.Operator.JoyBtnRaw);
IF bench.Operator.JoyBtnRaw AND NOT previousButton THEN buttonEdges := buttonEdges + 1; END_IF; previousButton := bench.Operator.JoyBtnRaw;
ASSERT_EQ(bench.Operator.JoyXRaw_ANA1, 5000, 'Pas de reprise apres OFF ON'); ASSERT_FALSE(bench.Operator.JoyBtnRaw, 'Bouton tenu ignore');
ADVANCE_TIME(10000000);
bench(RawPosM1 := raw1, RawPosM2 := raw2);
joy(RawX := bench.Operator.JoyXRaw_ANA1, RawY := bench.Operator.JoyYRaw_ANA2, RawButton := bench.Operator.JoyBtnRaw, Cfg := cfg, NeutralXMem := nx, NeutralYMem := ny);
home(DeadmanArmed := joy.DeadmanArmed, JoystickDeflected := NOT joy.AtNeutralXY, JoystickPull := joy.AxisCmdY.DirectionPositive, JoystickPush := joy.AxisCmdY.DirectionNegative, BtnValidation := bench.Operator.JoyBtnRaw);
IF bench.Operator.JoyBtnRaw AND NOT previousButton THEN buttonEdges := buttonEdges + 1; END_IF; previousButton := bench.Operator.JoyBtnRaw;
ASSERT_EQ(bench.Operator.JoyXRaw_ANA1, 5000, 'Pas de reprise apres OFF ON'); ASSERT_FALSE(bench.Operator.JoyBtnRaw, 'Bouton tenu ignore');
ADVANCE_TIME(10000000);
bench(RawPosM1 := raw1, RawPosM2 := raw2);
joy(RawX := bench.Operator.JoyXRaw_ANA1, RawY := bench.Operator.JoyYRaw_ANA2, RawButton := bench.Operator.JoyBtnRaw, Cfg := cfg, NeutralXMem := nx, NeutralYMem := ny);
home(DeadmanArmed := joy.DeadmanArmed, JoystickDeflected := NOT joy.AtNeutralXY, JoystickPull := joy.AxisCmdY.DirectionPositive, JoystickPush := joy.AxisCmdY.DirectionNegative, BtnValidation := bench.Operator.JoyBtnRaw);
IF bench.Operator.JoyBtnRaw AND NOT previousButton THEN buttonEdges := buttonEdges + 1; END_IF; previousButton := bench.Operator.JoyBtnRaw;
ASSERT_EQ(bench.Operator.JoyXRaw_ANA1, 5000, 'Pas de reprise apres OFF ON'); ASSERT_FALSE(bench.Operator.JoyBtnRaw, 'Bouton tenu ignore');
ADVANCE_TIME(10000000);
bench(RawPosM1 := raw1, RawPosM2 := raw2);
joy(RawX := bench.Operator.JoyXRaw_ANA1, RawY := bench.Operator.JoyYRaw_ANA2, RawButton := bench.Operator.JoyBtnRaw, Cfg := cfg, NeutralXMem := nx, NeutralYMem := ny);
home(DeadmanArmed := joy.DeadmanArmed, JoystickDeflected := NOT joy.AtNeutralXY, JoystickPull := joy.AxisCmdY.DirectionPositive, JoystickPush := joy.AxisCmdY.DirectionNegative, BtnValidation := bench.Operator.JoyBtnRaw);
IF bench.Operator.JoyBtnRaw AND NOT previousButton THEN buttonEdges := buttonEdges + 1; END_IF; previousButton := bench.Operator.JoyBtnRaw;
ASSERT_EQ(bench.Operator.JoyXRaw_ANA1, 5000, 'Pas de reprise apres OFF ON'); ASSERT_FALSE(bench.Operator.JoyBtnRaw, 'Bouton tenu ignore');
ADVANCE_TIME(10000000);
bench(RawPosM1 := raw1, RawPosM2 := raw2);
joy(RawX := bench.Operator.JoyXRaw_ANA1, RawY := bench.Operator.JoyYRaw_ANA2, RawButton := bench.Operator.JoyBtnRaw, Cfg := cfg, NeutralXMem := nx, NeutralYMem := ny);
home(DeadmanArmed := joy.DeadmanArmed, JoystickDeflected := NOT joy.AtNeutralXY, JoystickPull := joy.AxisCmdY.DirectionPositive, JoystickPush := joy.AxisCmdY.DirectionNegative, BtnValidation := bench.Operator.JoyBtnRaw);
IF bench.Operator.JoyBtnRaw AND NOT previousButton THEN buttonEdges := buttonEdges + 1; END_IF; previousButton := bench.Operator.JoyBtnRaw;
ASSERT_EQ(bench.Operator.JoyXRaw_ANA1, 5000, 'Pas de reprise apres OFF ON'); ASSERT_FALSE(bench.Operator.JoyBtnRaw, 'Bouton tenu ignore');
ADVANCE_TIME(10000000);
bench(RawPosM1 := raw1, RawPosM2 := raw2);
joy(RawX := bench.Operator.JoyXRaw_ANA1, RawY := bench.Operator.JoyYRaw_ANA2, RawButton := bench.Operator.JoyBtnRaw, Cfg := cfg, NeutralXMem := nx, NeutralYMem := ny);
home(DeadmanArmed := joy.DeadmanArmed, JoystickDeflected := NOT joy.AtNeutralXY, JoystickPull := joy.AxisCmdY.DirectionPositive, JoystickPush := joy.AxisCmdY.DirectionNegative, BtnValidation := bench.Operator.JoyBtnRaw);
IF bench.Operator.JoyBtnRaw AND NOT previousButton THEN buttonEdges := buttonEdges + 1; END_IF; previousButton := bench.Operator.JoyBtnRaw;
ASSERT_EQ(bench.Operator.JoyXRaw_ANA1, 5000, 'Pas de reprise apres OFF ON'); ASSERT_FALSE(bench.Operator.JoyBtnRaw, 'Bouton tenu ignore');
ADVANCE_TIME(10000000);
bench(RawPosM1 := raw1, RawPosM2 := raw2);
joy(RawX := bench.Operator.JoyXRaw_ANA1, RawY := bench.Operator.JoyYRaw_ANA2, RawButton := bench.Operator.JoyBtnRaw, Cfg := cfg, NeutralXMem := nx, NeutralYMem := ny);
home(DeadmanArmed := joy.DeadmanArmed, JoystickDeflected := NOT joy.AtNeutralXY, JoystickPull := joy.AxisCmdY.DirectionPositive, JoystickPush := joy.AxisCmdY.DirectionNegative, BtnValidation := bench.Operator.JoyBtnRaw);
IF bench.Operator.JoyBtnRaw AND NOT previousButton THEN buttonEdges := buttonEdges + 1; END_IF; previousButton := bench.Operator.JoyBtnRaw;
ASSERT_EQ(bench.Operator.JoyXRaw_ANA1, 5000, 'Pas de reprise apres OFF ON'); ASSERT_FALSE(bench.Operator.JoyBtnRaw, 'Bouton tenu ignore');
ADVANCE_TIME(10000000);
bench(RawPosM1 := raw1, RawPosM2 := raw2);
joy(RawX := bench.Operator.JoyXRaw_ANA1, RawY := bench.Operator.JoyYRaw_ANA2, RawButton := bench.Operator.JoyBtnRaw, Cfg := cfg, NeutralXMem := nx, NeutralYMem := ny);
home(DeadmanArmed := joy.DeadmanArmed, JoystickDeflected := NOT joy.AtNeutralXY, JoystickPull := joy.AxisCmdY.DirectionPositive, JoystickPush := joy.AxisCmdY.DirectionNegative, BtnValidation := bench.Operator.JoyBtnRaw);
IF bench.Operator.JoyBtnRaw AND NOT previousButton THEN buttonEdges := buttonEdges + 1; END_IF; previousButton := bench.Operator.JoyBtnRaw;
ASSERT_EQ(bench.Operator.JoyXRaw_ANA1, 5000, 'Pas de reprise apres OFF ON'); ASSERT_FALSE(bench.Operator.JoyBtnRaw, 'Bouton tenu ignore');
ADVANCE_TIME(10000000);
bench(RawPosM1 := raw1, RawPosM2 := raw2);
joy(RawX := bench.Operator.JoyXRaw_ANA1, RawY := bench.Operator.JoyYRaw_ANA2, RawButton := bench.Operator.JoyBtnRaw, Cfg := cfg, NeutralXMem := nx, NeutralYMem := ny);
home(DeadmanArmed := joy.DeadmanArmed, JoystickDeflected := NOT joy.AtNeutralXY, JoystickPull := joy.AxisCmdY.DirectionPositive, JoystickPush := joy.AxisCmdY.DirectionNegative, BtnValidation := bench.Operator.JoyBtnRaw);
IF bench.Operator.JoyBtnRaw AND NOT previousButton THEN buttonEdges := buttonEdges + 1; END_IF; previousButton := bench.Operator.JoyBtnRaw;
ASSERT_EQ(bench.Operator.JoyXRaw_ANA1, 5000, 'Pas de reprise apres OFF ON'); ASSERT_FALSE(bench.Operator.JoyBtnRaw, 'Bouton tenu ignore');
ADVANCE_TIME(10000000);
bench(RawPosM1 := raw1, RawPosM2 := raw2);
joy(RawX := bench.Operator.JoyXRaw_ANA1, RawY := bench.Operator.JoyYRaw_ANA2, RawButton := bench.Operator.JoyBtnRaw, Cfg := cfg, NeutralXMem := nx, NeutralYMem := ny);
home(DeadmanArmed := joy.DeadmanArmed, JoystickDeflected := NOT joy.AtNeutralXY, JoystickPull := joy.AxisCmdY.DirectionPositive, JoystickPush := joy.AxisCmdY.DirectionNegative, BtnValidation := bench.Operator.JoyBtnRaw);
IF bench.Operator.JoyBtnRaw AND NOT previousButton THEN buttonEdges := buttonEdges + 1; END_IF; previousButton := bench.Operator.JoyBtnRaw;
ASSERT_EQ(bench.Operator.JoyXRaw_ANA1, 5000, 'Pas de reprise apres OFF ON'); ASSERT_FALSE(bench.Operator.JoyBtnRaw, 'Bouton tenu ignore');
ADVANCE_TIME(10000000);
bench(RawPosM1 := raw1, RawPosM2 := raw2);
joy(RawX := bench.Operator.JoyXRaw_ANA1, RawY := bench.Operator.JoyYRaw_ANA2, RawButton := bench.Operator.JoyBtnRaw, Cfg := cfg, NeutralXMem := nx, NeutralYMem := ny);
home(DeadmanArmed := joy.DeadmanArmed, JoystickDeflected := NOT joy.AtNeutralXY, JoystickPull := joy.AxisCmdY.DirectionPositive, JoystickPush := joy.AxisCmdY.DirectionNegative, BtnValidation := bench.Operator.JoyBtnRaw);
IF bench.Operator.JoyBtnRaw AND NOT previousButton THEN buttonEdges := buttonEdges + 1; END_IF; previousButton := bench.Operator.JoyBtnRaw;
ASSERT_EQ(bench.Operator.JoyXRaw_ANA1, 5000, 'Pas de reprise apres OFF ON'); ASSERT_FALSE(bench.Operator.JoyBtnRaw, 'Bouton tenu ignore');
ADVANCE_TIME(10000000);
bench(RawPosM1 := raw1, RawPosM2 := raw2);
joy(RawX := bench.Operator.JoyXRaw_ANA1, RawY := bench.Operator.JoyYRaw_ANA2, RawButton := bench.Operator.JoyBtnRaw, Cfg := cfg, NeutralXMem := nx, NeutralYMem := ny);
home(DeadmanArmed := joy.DeadmanArmed, JoystickDeflected := NOT joy.AtNeutralXY, JoystickPull := joy.AxisCmdY.DirectionPositive, JoystickPush := joy.AxisCmdY.DirectionNegative, BtnValidation := bench.Operator.JoyBtnRaw);
IF bench.Operator.JoyBtnRaw AND NOT previousButton THEN buttonEdges := buttonEdges + 1; END_IF; previousButton := bench.Operator.JoyBtnRaw;
ASSERT_EQ(bench.Operator.JoyXRaw_ANA1, 5000, 'Pas de reprise apres OFF ON'); ASSERT_FALSE(bench.Operator.JoyBtnRaw, 'Bouton tenu ignore');
ADVANCE_TIME(10000000);
bench(RawPosM1 := raw1, RawPosM2 := raw2);
joy(RawX := bench.Operator.JoyXRaw_ANA1, RawY := bench.Operator.JoyYRaw_ANA2, RawButton := bench.Operator.JoyBtnRaw, Cfg := cfg, NeutralXMem := nx, NeutralYMem := ny);
home(DeadmanArmed := joy.DeadmanArmed, JoystickDeflected := NOT joy.AtNeutralXY, JoystickPull := joy.AxisCmdY.DirectionPositive, JoystickPush := joy.AxisCmdY.DirectionNegative, BtnValidation := bench.Operator.JoyBtnRaw);
IF bench.Operator.JoyBtnRaw AND NOT previousButton THEN buttonEdges := buttonEdges + 1; END_IF; previousButton := bench.Operator.JoyBtnRaw;
ASSERT_EQ(bench.Operator.JoyXRaw_ANA1, 5000, 'Pas de reprise apres OFF ON'); ASSERT_FALSE(bench.Operator.JoyBtnRaw, 'Bouton tenu ignore');
ADVANCE_TIME(10000000);
bench(RawPosM1 := raw1, RawPosM2 := raw2);
joy(RawX := bench.Operator.JoyXRaw_ANA1, RawY := bench.Operator.JoyYRaw_ANA2, RawButton := bench.Operator.JoyBtnRaw, Cfg := cfg, NeutralXMem := nx, NeutralYMem := ny);
home(DeadmanArmed := joy.DeadmanArmed, JoystickDeflected := NOT joy.AtNeutralXY, JoystickPull := joy.AxisCmdY.DirectionPositive, JoystickPush := joy.AxisCmdY.DirectionNegative, BtnValidation := bench.Operator.JoyBtnRaw);
IF bench.Operator.JoyBtnRaw AND NOT previousButton THEN buttonEdges := buttonEdges + 1; END_IF; previousButton := bench.Operator.JoyBtnRaw;
ASSERT_EQ(bench.Operator.JoyXRaw_ANA1, 5000, 'Pas de reprise apres OFF ON'); ASSERT_FALSE(bench.Operator.JoyBtnRaw, 'Bouton tenu ignore');
ADVANCE_TIME(10000000);
bench(RawPosM1 := raw1, RawPosM2 := raw2);
joy(RawX := bench.Operator.JoyXRaw_ANA1, RawY := bench.Operator.JoyYRaw_ANA2, RawButton := bench.Operator.JoyBtnRaw, Cfg := cfg, NeutralXMem := nx, NeutralYMem := ny);
home(DeadmanArmed := joy.DeadmanArmed, JoystickDeflected := NOT joy.AtNeutralXY, JoystickPull := joy.AxisCmdY.DirectionPositive, JoystickPush := joy.AxisCmdY.DirectionNegative, BtnValidation := bench.Operator.JoyBtnRaw);
IF bench.Operator.JoyBtnRaw AND NOT previousButton THEN buttonEdges := buttonEdges + 1; END_IF; previousButton := bench.Operator.JoyBtnRaw;
ASSERT_EQ(bench.Operator.JoyXRaw_ANA1, 5000, 'Pas de reprise apres OFF ON'); ASSERT_FALSE(bench.Operator.JoyBtnRaw, 'Bouton tenu ignore');
ADVANCE_TIME(10000000);
bench(RawPosM1 := raw1, RawPosM2 := raw2);
joy(RawX := bench.Operator.JoyXRaw_ANA1, RawY := bench.Operator.JoyYRaw_ANA2, RawButton := bench.Operator.JoyBtnRaw, Cfg := cfg, NeutralXMem := nx, NeutralYMem := ny);
home(DeadmanArmed := joy.DeadmanArmed, JoystickDeflected := NOT joy.AtNeutralXY, JoystickPull := joy.AxisCmdY.DirectionPositive, JoystickPush := joy.AxisCmdY.DirectionNegative, BtnValidation := bench.Operator.JoyBtnRaw);
IF bench.Operator.JoyBtnRaw AND NOT previousButton THEN buttonEdges := buttonEdges + 1; END_IF; previousButton := bench.Operator.JoyBtnRaw;
ASSERT_EQ(bench.Operator.JoyXRaw_ANA1, 5000, 'Pas de reprise apres OFF ON'); ASSERT_FALSE(bench.Operator.JoyBtnRaw, 'Bouton tenu ignore');
ADVANCE_TIME(10000000);
bench(RawPosM1 := raw1, RawPosM2 := raw2);
joy(RawX := bench.Operator.JoyXRaw_ANA1, RawY := bench.Operator.JoyYRaw_ANA2, RawButton := bench.Operator.JoyBtnRaw, Cfg := cfg, NeutralXMem := nx, NeutralYMem := ny);
home(DeadmanArmed := joy.DeadmanArmed, JoystickDeflected := NOT joy.AtNeutralXY, JoystickPull := joy.AxisCmdY.DirectionPositive, JoystickPush := joy.AxisCmdY.DirectionNegative, BtnValidation := bench.Operator.JoyBtnRaw);
IF bench.Operator.JoyBtnRaw AND NOT previousButton THEN buttonEdges := buttonEdges + 1; END_IF; previousButton := bench.Operator.JoyBtnRaw;
ASSERT_EQ(bench.Operator.JoyXRaw_ANA1, 5000, 'Pas de reprise apres OFF ON'); ASSERT_FALSE(bench.Operator.JoyBtnRaw, 'Bouton tenu ignore');
ADVANCE_TIME(10000000);
bench(RawPosM1 := raw1, RawPosM2 := raw2);
joy(RawX := bench.Operator.JoyXRaw_ANA1, RawY := bench.Operator.JoyYRaw_ANA2, RawButton := bench.Operator.JoyBtnRaw, Cfg := cfg, NeutralXMem := nx, NeutralYMem := ny);
home(DeadmanArmed := joy.DeadmanArmed, JoystickDeflected := NOT joy.AtNeutralXY, JoystickPull := joy.AxisCmdY.DirectionPositive, JoystickPush := joy.AxisCmdY.DirectionNegative, BtnValidation := bench.Operator.JoyBtnRaw);
IF bench.Operator.JoyBtnRaw AND NOT previousButton THEN buttonEdges := buttonEdges + 1; END_IF; previousButton := bench.Operator.JoyBtnRaw;
ASSERT_EQ(bench.Operator.JoyXRaw_ANA1, 5000, 'Pas de reprise apres OFF ON'); ASSERT_FALSE(bench.Operator.JoyBtnRaw, 'Bouton tenu ignore');
ADVANCE_TIME(10000000);
bench(RawPosM1 := raw1, RawPosM2 := raw2);
joy(RawX := bench.Operator.JoyXRaw_ANA1, RawY := bench.Operator.JoyYRaw_ANA2, RawButton := bench.Operator.JoyBtnRaw, Cfg := cfg, NeutralXMem := nx, NeutralYMem := ny);
home(DeadmanArmed := joy.DeadmanArmed, JoystickDeflected := NOT joy.AtNeutralXY, JoystickPull := joy.AxisCmdY.DirectionPositive, JoystickPush := joy.AxisCmdY.DirectionNegative, BtnValidation := bench.Operator.JoyBtnRaw);
IF bench.Operator.JoyBtnRaw AND NOT previousButton THEN buttonEdges := buttonEdges + 1; END_IF; previousButton := bench.Operator.JoyBtnRaw;
ASSERT_EQ(bench.Operator.JoyXRaw_ANA1, 5000, 'Pas de reprise apres OFF ON'); ASSERT_FALSE(bench.Operator.JoyBtnRaw, 'Bouton tenu ignore');
ADVANCE_TIME(10000000);
bench(RawPosM1 := raw1, RawPosM2 := raw2);
joy(RawX := bench.Operator.JoyXRaw_ANA1, RawY := bench.Operator.JoyYRaw_ANA2, RawButton := bench.Operator.JoyBtnRaw, Cfg := cfg, NeutralXMem := nx, NeutralYMem := ny);
home(DeadmanArmed := joy.DeadmanArmed, JoystickDeflected := NOT joy.AtNeutralXY, JoystickPull := joy.AxisCmdY.DirectionPositive, JoystickPush := joy.AxisCmdY.DirectionNegative, BtnValidation := bench.Operator.JoyBtnRaw);
IF bench.Operator.JoyBtnRaw AND NOT previousButton THEN buttonEdges := buttonEdges + 1; END_IF; previousButton := bench.Operator.JoyBtnRaw;
ASSERT_EQ(bench.Operator.JoyXRaw_ANA1, 5000, 'Pas de reprise apres OFF ON'); ASSERT_FALSE(bench.Operator.JoyBtnRaw, 'Bouton tenu ignore');
ADVANCE_TIME(10000000);
bench(RawPosM1 := raw1, RawPosM2 := raw2);
joy(RawX := bench.Operator.JoyXRaw_ANA1, RawY := bench.Operator.JoyYRaw_ANA2, RawButton := bench.Operator.JoyBtnRaw, Cfg := cfg, NeutralXMem := nx, NeutralYMem := ny);
home(DeadmanArmed := joy.DeadmanArmed, JoystickDeflected := NOT joy.AtNeutralXY, JoystickPull := joy.AxisCmdY.DirectionPositive, JoystickPush := joy.AxisCmdY.DirectionNegative, BtnValidation := bench.Operator.JoyBtnRaw);
IF bench.Operator.JoyBtnRaw AND NOT previousButton THEN buttonEdges := buttonEdges + 1; END_IF; previousButton := bench.Operator.JoyBtnRaw;
ASSERT_EQ(bench.Operator.JoyXRaw_ANA1, 5000, 'Pas de reprise apres OFF ON'); ASSERT_FALSE(bench.Operator.JoyBtnRaw, 'Bouton tenu ignore');
ADVANCE_TIME(10000000);
bench(RawPosM1 := raw1, RawPosM2 := raw2);
joy(RawX := bench.Operator.JoyXRaw_ANA1, RawY := bench.Operator.JoyYRaw_ANA2, RawButton := bench.Operator.JoyBtnRaw, Cfg := cfg, NeutralXMem := nx, NeutralYMem := ny);
home(DeadmanArmed := joy.DeadmanArmed, JoystickDeflected := NOT joy.AtNeutralXY, JoystickPull := joy.AxisCmdY.DirectionPositive, JoystickPush := joy.AxisCmdY.DirectionNegative, BtnValidation := bench.Operator.JoyBtnRaw);
IF bench.Operator.JoyBtnRaw AND NOT previousButton THEN buttonEdges := buttonEdges + 1; END_IF; previousButton := bench.Operator.JoyBtnRaw;
ASSERT_EQ(bench.Operator.JoyXRaw_ANA1, 5000, 'Pas de reprise apres OFF ON'); ASSERT_FALSE(bench.Operator.JoyBtnRaw, 'Bouton tenu ignore');
ADVANCE_TIME(10000000);
bench(RawPosM1 := raw1, RawPosM2 := raw2);
joy(RawX := bench.Operator.JoyXRaw_ANA1, RawY := bench.Operator.JoyYRaw_ANA2, RawButton := bench.Operator.JoyBtnRaw, Cfg := cfg, NeutralXMem := nx, NeutralYMem := ny);
home(DeadmanArmed := joy.DeadmanArmed, JoystickDeflected := NOT joy.AtNeutralXY, JoystickPull := joy.AxisCmdY.DirectionPositive, JoystickPush := joy.AxisCmdY.DirectionNegative, BtnValidation := bench.Operator.JoyBtnRaw);
IF bench.Operator.JoyBtnRaw AND NOT previousButton THEN buttonEdges := buttonEdges + 1; END_IF; previousButton := bench.Operator.JoyBtnRaw;
ASSERT_EQ(bench.Operator.JoyXRaw_ANA1, 5000, 'Pas de reprise apres OFF ON'); ASSERT_FALSE(bench.Operator.JoyBtnRaw, 'Bouton tenu ignore');
ADVANCE_TIME(10000000);
bench(RawPosM1 := raw1, RawPosM2 := raw2);
joy(RawX := bench.Operator.JoyXRaw_ANA1, RawY := bench.Operator.JoyYRaw_ANA2, RawButton := bench.Operator.JoyBtnRaw, Cfg := cfg, NeutralXMem := nx, NeutralYMem := ny);
home(DeadmanArmed := joy.DeadmanArmed, JoystickDeflected := NOT joy.AtNeutralXY, JoystickPull := joy.AxisCmdY.DirectionPositive, JoystickPush := joy.AxisCmdY.DirectionNegative, BtnValidation := bench.Operator.JoyBtnRaw);
IF bench.Operator.JoyBtnRaw AND NOT previousButton THEN buttonEdges := buttonEdges + 1; END_IF; previousButton := bench.Operator.JoyBtnRaw;
ASSERT_EQ(bench.Operator.JoyXRaw_ANA1, 5000, 'Pas de reprise apres OFF ON'); ASSERT_FALSE(bench.Operator.JoyBtnRaw, 'Bouton tenu ignore');
ADVANCE_TIME(10000000);
bench(RawPosM1 := raw1, RawPosM2 := raw2);
joy(RawX := bench.Operator.JoyXRaw_ANA1, RawY := bench.Operator.JoyYRaw_ANA2, RawButton := bench.Operator.JoyBtnRaw, Cfg := cfg, NeutralXMem := nx, NeutralYMem := ny);
home(DeadmanArmed := joy.DeadmanArmed, JoystickDeflected := NOT joy.AtNeutralXY, JoystickPull := joy.AxisCmdY.DirectionPositive, JoystickPush := joy.AxisCmdY.DirectionNegative, BtnValidation := bench.Operator.JoyBtnRaw);
IF bench.Operator.JoyBtnRaw AND NOT previousButton THEN buttonEdges := buttonEdges + 1; END_IF; previousButton := bench.Operator.JoyBtnRaw;
ASSERT_EQ(bench.Operator.JoyXRaw_ANA1, 5000, 'Pas de reprise apres OFF ON'); ASSERT_FALSE(bench.Operator.JoyBtnRaw, 'Bouton tenu ignore');
ADVANCE_TIME(10000000);
bench(RawPosM1 := raw1, RawPosM2 := raw2);
joy(RawX := bench.Operator.JoyXRaw_ANA1, RawY := bench.Operator.JoyYRaw_ANA2, RawButton := bench.Operator.JoyBtnRaw, Cfg := cfg, NeutralXMem := nx, NeutralYMem := ny);
home(DeadmanArmed := joy.DeadmanArmed, JoystickDeflected := NOT joy.AtNeutralXY, JoystickPull := joy.AxisCmdY.DirectionPositive, JoystickPush := joy.AxisCmdY.DirectionNegative, BtnValidation := bench.Operator.JoyBtnRaw);
IF bench.Operator.JoyBtnRaw AND NOT previousButton THEN buttonEdges := buttonEdges + 1; END_IF; previousButton := bench.Operator.JoyBtnRaw;
ASSERT_EQ(bench.Operator.JoyXRaw_ANA1, 5000, 'Pas de reprise apres OFF ON'); ASSERT_FALSE(bench.Operator.JoyBtnRaw, 'Bouton tenu ignore');
ADVANCE_TIME(10000000);
bench(RawPosM1 := raw1, RawPosM2 := raw2);
joy(RawX := bench.Operator.JoyXRaw_ANA1, RawY := bench.Operator.JoyYRaw_ANA2, RawButton := bench.Operator.JoyBtnRaw, Cfg := cfg, NeutralXMem := nx, NeutralYMem := ny);
home(DeadmanArmed := joy.DeadmanArmed, JoystickDeflected := NOT joy.AtNeutralXY, JoystickPull := joy.AxisCmdY.DirectionPositive, JoystickPush := joy.AxisCmdY.DirectionNegative, BtnValidation := bench.Operator.JoyBtnRaw);
IF bench.Operator.JoyBtnRaw AND NOT previousButton THEN buttonEdges := buttonEdges + 1; END_IF; previousButton := bench.Operator.JoyBtnRaw;
ASSERT_EQ(bench.Operator.JoyXRaw_ANA1, 5000, 'Pas de reprise apres OFF ON'); ASSERT_FALSE(bench.Operator.JoyBtnRaw, 'Bouton tenu ignore');
ADVANCE_TIME(10000000);
bench(RawPosM1 := raw1, RawPosM2 := raw2);
joy(RawX := bench.Operator.JoyXRaw_ANA1, RawY := bench.Operator.JoyYRaw_ANA2, RawButton := bench.Operator.JoyBtnRaw, Cfg := cfg, NeutralXMem := nx, NeutralYMem := ny);
home(DeadmanArmed := joy.DeadmanArmed, JoystickDeflected := NOT joy.AtNeutralXY, JoystickPull := joy.AxisCmdY.DirectionPositive, JoystickPush := joy.AxisCmdY.DirectionNegative, BtnValidation := bench.Operator.JoyBtnRaw);
IF bench.Operator.JoyBtnRaw AND NOT previousButton THEN buttonEdges := buttonEdges + 1; END_IF; previousButton := bench.Operator.JoyBtnRaw;
ASSERT_EQ(bench.Operator.JoyXRaw_ANA1, 5000, 'Pas de reprise apres OFF ON'); ASSERT_FALSE(bench.Operator.JoyBtnRaw, 'Bouton tenu ignore');
ADVANCE_TIME(10000000);
bench(RawPosM1 := raw1, RawPosM2 := raw2);
joy(RawX := bench.Operator.JoyXRaw_ANA1, RawY := bench.Operator.JoyYRaw_ANA2, RawButton := bench.Operator.JoyBtnRaw, Cfg := cfg, NeutralXMem := nx, NeutralYMem := ny);
home(DeadmanArmed := joy.DeadmanArmed, JoystickDeflected := NOT joy.AtNeutralXY, JoystickPull := joy.AxisCmdY.DirectionPositive, JoystickPush := joy.AxisCmdY.DirectionNegative, BtnValidation := bench.Operator.JoyBtnRaw);
IF bench.Operator.JoyBtnRaw AND NOT previousButton THEN buttonEdges := buttonEdges + 1; END_IF; previousButton := bench.Operator.JoyBtnRaw;
ASSERT_EQ(bench.Operator.JoyXRaw_ANA1, 5000, 'Pas de reprise apres OFF ON'); ASSERT_FALSE(bench.Operator.JoyBtnRaw, 'Bouton tenu ignore');
ADVANCE_TIME(10000000);
bench(RawPosM1 := raw1, RawPosM2 := raw2);
joy(RawX := bench.Operator.JoyXRaw_ANA1, RawY := bench.Operator.JoyYRaw_ANA2, RawButton := bench.Operator.JoyBtnRaw, Cfg := cfg, NeutralXMem := nx, NeutralYMem := ny);
home(DeadmanArmed := joy.DeadmanArmed, JoystickDeflected := NOT joy.AtNeutralXY, JoystickPull := joy.AxisCmdY.DirectionPositive, JoystickPush := joy.AxisCmdY.DirectionNegative, BtnValidation := bench.Operator.JoyBtnRaw);
IF bench.Operator.JoyBtnRaw AND NOT previousButton THEN buttonEdges := buttonEdges + 1; END_IF; previousButton := bench.Operator.JoyBtnRaw;
ASSERT_EQ(bench.Operator.JoyXRaw_ANA1, 5000, 'Pas de reprise apres OFF ON'); ASSERT_FALSE(bench.Operator.JoyBtnRaw, 'Bouton tenu ignore');
ADVANCE_TIME(10000000);
bench(RawPosM1 := raw1, RawPosM2 := raw2);
joy(RawX := bench.Operator.JoyXRaw_ANA1, RawY := bench.Operator.JoyYRaw_ANA2, RawButton := bench.Operator.JoyBtnRaw, Cfg := cfg, NeutralXMem := nx, NeutralYMem := ny);
home(DeadmanArmed := joy.DeadmanArmed, JoystickDeflected := NOT joy.AtNeutralXY, JoystickPull := joy.AxisCmdY.DirectionPositive, JoystickPush := joy.AxisCmdY.DirectionNegative, BtnValidation := bench.Operator.JoyBtnRaw);
IF bench.Operator.JoyBtnRaw AND NOT previousButton THEN buttonEdges := buttonEdges + 1; END_IF; previousButton := bench.Operator.JoyBtnRaw;
ASSERT_EQ(bench.Operator.JoyXRaw_ANA1, 5000, 'Pas de reprise apres OFF ON'); ASSERT_FALSE(bench.Operator.JoyBtnRaw, 'Bouton tenu ignore');
ADVANCE_TIME(10000000);
bench(RawPosM1 := raw1, RawPosM2 := raw2);
joy(RawX := bench.Operator.JoyXRaw_ANA1, RawY := bench.Operator.JoyYRaw_ANA2, RawButton := bench.Operator.JoyBtnRaw, Cfg := cfg, NeutralXMem := nx, NeutralYMem := ny);
home(DeadmanArmed := joy.DeadmanArmed, JoystickDeflected := NOT joy.AtNeutralXY, JoystickPull := joy.AxisCmdY.DirectionPositive, JoystickPush := joy.AxisCmdY.DirectionNegative, BtnValidation := bench.Operator.JoyBtnRaw);
IF bench.Operator.JoyBtnRaw AND NOT previousButton THEN buttonEdges := buttonEdges + 1; END_IF; previousButton := bench.Operator.JoyBtnRaw;
ASSERT_EQ(bench.Operator.JoyXRaw_ANA1, 5000, 'Pas de reprise apres OFF ON'); ASSERT_FALSE(bench.Operator.JoyBtnRaw, 'Bouton tenu ignore');
ADVANCE_TIME(10000000);
bench(RawPosM1 := raw1, RawPosM2 := raw2);
joy(RawX := bench.Operator.JoyXRaw_ANA1, RawY := bench.Operator.JoyYRaw_ANA2, RawButton := bench.Operator.JoyBtnRaw, Cfg := cfg, NeutralXMem := nx, NeutralYMem := ny);
home(DeadmanArmed := joy.DeadmanArmed, JoystickDeflected := NOT joy.AtNeutralXY, JoystickPull := joy.AxisCmdY.DirectionPositive, JoystickPush := joy.AxisCmdY.DirectionNegative, BtnValidation := bench.Operator.JoyBtnRaw);
IF bench.Operator.JoyBtnRaw AND NOT previousButton THEN buttonEdges := buttonEdges + 1; END_IF; previousButton := bench.Operator.JoyBtnRaw;
ASSERT_EQ(bench.Operator.JoyXRaw_ANA1, 5000, 'Pas de reprise apres OFF ON'); ASSERT_FALSE(bench.Operator.JoyBtnRaw, 'Bouton tenu ignore');
ADVANCE_TIME(10000000);
bench(RawPosM1 := raw1, RawPosM2 := raw2);
joy(RawX := bench.Operator.JoyXRaw_ANA1, RawY := bench.Operator.JoyYRaw_ANA2, RawButton := bench.Operator.JoyBtnRaw, Cfg := cfg, NeutralXMem := nx, NeutralYMem := ny);
home(DeadmanArmed := joy.DeadmanArmed, JoystickDeflected := NOT joy.AtNeutralXY, JoystickPull := joy.AxisCmdY.DirectionPositive, JoystickPush := joy.AxisCmdY.DirectionNegative, BtnValidation := bench.Operator.JoyBtnRaw);
IF bench.Operator.JoyBtnRaw AND NOT previousButton THEN buttonEdges := buttonEdges + 1; END_IF; previousButton := bench.Operator.JoyBtnRaw;
ASSERT_EQ(bench.Operator.JoyXRaw_ANA1, 5000, 'Pas de reprise apres OFF ON'); ASSERT_FALSE(bench.Operator.JoyBtnRaw, 'Bouton tenu ignore');
ADVANCE_TIME(10000000);
bench(RawPosM1 := raw1, RawPosM2 := raw2);
joy(RawX := bench.Operator.JoyXRaw_ANA1, RawY := bench.Operator.JoyYRaw_ANA2, RawButton := bench.Operator.JoyBtnRaw, Cfg := cfg, NeutralXMem := nx, NeutralYMem := ny);
home(DeadmanArmed := joy.DeadmanArmed, JoystickDeflected := NOT joy.AtNeutralXY, JoystickPull := joy.AxisCmdY.DirectionPositive, JoystickPush := joy.AxisCmdY.DirectionNegative, BtnValidation := bench.Operator.JoyBtnRaw);
IF bench.Operator.JoyBtnRaw AND NOT previousButton THEN buttonEdges := buttonEdges + 1; END_IF; previousButton := bench.Operator.JoyBtnRaw;
ASSERT_EQ(bench.Operator.JoyXRaw_ANA1, 5000, 'Pas de reprise apres OFF ON'); ASSERT_FALSE(bench.Operator.JoyBtnRaw, 'Bouton tenu ignore');
ADVANCE_TIME(10000000);
bench(RawPosM1 := raw1, RawPosM2 := raw2);
joy(RawX := bench.Operator.JoyXRaw_ANA1, RawY := bench.Operator.JoyYRaw_ANA2, RawButton := bench.Operator.JoyBtnRaw, Cfg := cfg, NeutralXMem := nx, NeutralYMem := ny);
home(DeadmanArmed := joy.DeadmanArmed, JoystickDeflected := NOT joy.AtNeutralXY, JoystickPull := joy.AxisCmdY.DirectionPositive, JoystickPush := joy.AxisCmdY.DirectionNegative, BtnValidation := bench.Operator.JoyBtnRaw);
IF bench.Operator.JoyBtnRaw AND NOT previousButton THEN buttonEdges := buttonEdges + 1; END_IF; previousButton := bench.Operator.JoyBtnRaw;
ASSERT_EQ(bench.Operator.JoyXRaw_ANA1, 5000, 'Pas de reprise apres OFF ON'); ASSERT_FALSE(bench.Operator.JoyBtnRaw, 'Bouton tenu ignore');
ADVANCE_TIME(10000000);
bench(RawPosM1 := raw1, RawPosM2 := raw2);
joy(RawX := bench.Operator.JoyXRaw_ANA1, RawY := bench.Operator.JoyYRaw_ANA2, RawButton := bench.Operator.JoyBtnRaw, Cfg := cfg, NeutralXMem := nx, NeutralYMem := ny);
home(DeadmanArmed := joy.DeadmanArmed, JoystickDeflected := NOT joy.AtNeutralXY, JoystickPull := joy.AxisCmdY.DirectionPositive, JoystickPush := joy.AxisCmdY.DirectionNegative, BtnValidation := bench.Operator.JoyBtnRaw);
IF bench.Operator.JoyBtnRaw AND NOT previousButton THEN buttonEdges := buttonEdges + 1; END_IF; previousButton := bench.Operator.JoyBtnRaw;
ASSERT_EQ(bench.Operator.JoyXRaw_ANA1, 5000, 'Pas de reprise apres OFF ON'); ASSERT_FALSE(bench.Operator.JoyBtnRaw, 'Bouton tenu ignore');
END_TEST
